(* Logix 5000 project; controller TFF vendor 1 type 14 code 107 rev 34.11; software revision 34.03; part 5 of 36 *)

        [11].DelayTimerSP := 1, [11].ActiveStateCFg := 1, [11].RealInputCfg := 1, [11].InputAddressCfg := 11, [12].Tag := 'XS012', [12].DelayTimer.PRE := 1000, [12].DelayTimerSP := 1, [12].EnableCfg := 1, [12].ActiveStateCFg := 1, [12].RealInputCfg := 1, [12].InputAddressCfg := 12, [13].Tag := 'XC102_3DF', [13].AlarmCurrentValue := 1, [13].Override := 1, [13].DelayTimer.PRE := 1000, [13].DelayTimer.ACC := 1007, [13].DelayTimer.EN := 1, [13].DelayTimer.DN := 1, [13].DelayTimerSP := 1, [13].Priority := 1, [13].EnableCfg := 1, [13].ActiveStateCFg := 1, [13].RealInputCfg := 1, [13].InputAddressCfg := 13, [13].AlarmCfg := 1, [13].OverrideCfg := 1, [13].PriorityCfg := 1, [14].Tag := 'SIC003DF', [14].AlarmCurrentValue := 1, [14].Override := 1, [14].DelayTimer.PRE := 1000, [14].DelayTimer.ACC := 1005, [14].DelayTimer.EN := 1, [14].DelayTimer.DN := 1, [14].DelayTimerSP := 1, [14].Priority := 1, [14].EnableCfg := 1, [14].ActiveStateCFg := 1, [14].RealInputCfg := 1, [14].InputAddressCfg := 14, [14].AlarmCfg := 1, [14].OverrideCfg := 1, [14].PriorityCfg := 1, [15].Tag := 'SRL001', [15].SoftInput := 1, [15].DelayTimer.PRE := 2000, [15].DelayTimerSP := 2, [15].EnableCfg := 1, [15].ActiveStateCFg := 1, [15].RealInputCfg := 1, [15].InputAddressCfg := 15, [16].AlarmCurrentValue := 1, [16].Override := 1, [16].SoftInput := 1, [16].DelayTimer.PRE := 1000, [16].DelayTimer.ACC := 1018, [16].DelayTimer.EN := 1, [16].DelayTimer.DN := 1, [16].DelayTimerSP := 1, [16].Priority := 1,
        [16].ActiveStateCFg := 1, [16].RealInputCfg := 1, [16].InputAddressCfg := 16, [16].OverrideCfg := 1, [16].PriorityCfg := 1, [17].AlarmCurrentValue := 1, [17].Override := 1, [17].SoftInput := 1, [17].DelayTimer.PRE := 1000, [17].DelayTimer.ACC := 1018, [17].DelayTimer.EN := 1, [17].DelayTimer.DN := 1, [17].DelayTimerSP := 1, [17].Priority := 1, [17].ActiveStateCFg := 1, [17].RealInputCfg := 1, [17].InputAddressCfg := 17, [17].OverrideCfg := 1, [17].PriorityCfg := 1, [18].AlarmCurrentValue := 1, [18].Override := 1, [18].DelayTimer.PRE := 1000, [18].DelayTimer.ACC := 1018, [18].DelayTimer.EN := 1, [18].DelayTimer.DN := 1, [18].DelayTimerSP := 1, [18].Priority := 1, [18].ActiveStateCFg := 1, [18].RealInputCfg := 1, [18].InputAddressCfg := 18, [18].OverrideCfg := 1, [18].PriorityCfg := 1, [19].AlarmCurrentValue := 1, [19].Override := 1, [19].DelayTimer.PRE := 1000, [19].DelayTimer.ACC := 1019, [19].DelayTimer.EN := 1, [19].DelayTimer.DN := 1, [19].DelayTimerSP := 1, [19].ActiveStateCFg := 1, [19].RealInputCfg := 1, [19].InputAddressCfg := 19, [19].OverrideCfg := 1, [19].PriorityCfg := 1, [20].AlarmCurrentValue := 1, [20].Override := 1, [20].DelayTimer.PRE := 1000, [20].DelayTimer.ACC := 1019, [20].DelayTimer.EN := 1, [20].DelayTimer.DN := 1, [20].DelayTimerSP := 1, [20].ActiveStateCFg := 1, [20].RealInputCfg := 1, [20].InputAddressCfg := 20, [20].OverrideCfg := 1, [20].PriorityCfg := 1, [21].AlarmCurrentValue := 1, [21].AlarmAck := 1, [21].Alarm := 1, [21].Mimic := 5,
        [21].DelayTimer.PRE := 1000, [21].DelayTimer.ACC := 1003, [21].DelayTimer.EN := 1, [21].DelayTimer.DN := 1, [21].DelayTimerSP := 1, [21].Priority := 1, [21].ActiveStateCFg := 1, [21].RealInputCfg := 1, [21].InputAddressCfg := 21, [21].AlarmONS := 1, [22].AlarmCurrentValue := 1, [22].AlarmAck := 1, [22].Alarm := 1, [22].Mimic := 5, [22].DelayTimer.PRE := 1000, [22].DelayTimer.ACC := 1004, [22].DelayTimer.EN := 1, [22].DelayTimer.DN := 1, [22].DelayTimerSP := 1, [22].Priority := 1, [22].ActiveStateCFg := 1, [22].RealInputCfg := 1, [22].InputAddressCfg := 22, [22].AlarmONS := 1, [23].AlarmCurrentValue := 1, [23].Override := 1, [23].DelayTimer.PRE := 1000, [23].DelayTimer.ACC := 1018, [23].DelayTimer.EN := 1, [23].DelayTimer.DN := 1, [23].DelayTimerSP := 1, [23].Priority := 1, [23].ActiveStateCFg := 1, [23].RealInputCfg := 1, [23].InputAddressCfg := 23, [23].OverrideCfg := 1, [23].PriorityCfg := 1, [24].AlarmCurrentValue := 1, [24].Override := 1, [24].DelayTimer.PRE := 1000, [24].DelayTimer.ACC := 1018, [24].DelayTimer.EN := 1, [24].DelayTimer.DN := 1, [24].DelayTimerSP := 1, [24].Priority := 1, [24].ActiveStateCFg := 1, [24].RealInputCfg := 1, [24].InputAddressCfg := 24, [24].OverrideCfg := 1, [24].PriorityCfg := 1, [25].AlarmCurrentValue := 1, [25].Override := 1, [25].DelayTimer.PRE := 20000, [25].DelayTimerSP := 2, [25].Priority := 1, [25].ActiveStateCFg := 1, [25].RealInputCfg := 1, [25].InputAddressCfg := 25, [25].OverrideCfg := 1, [25].PriorityCfg := 1,
        [25].Cond1Cfg := 1, [27].SoftInput := 1, [28].SoftInput := 1, [29].SoftInput := 1, [30].SoftInput := 1, [34].Tag := 'DI1', [34].Override := 1, [34].SoftInput := 1, [34].ActiveStateCFg := 1, [34].RealInputCfg := 1, [34].InputAddressCfg := 34, [34].OverrideCfg := 1, [34].PriorityCfg := 1, [35].Tag := 'DI2', [35].Override := 1, [35].ActiveStateCFg := 1, [35].RealInputCfg := 1, [35].InputAddressCfg := 35, [35].OverrideCfg := 1, [35].PriorityCfg := 1, [36].Tag := 'DI3', [36].Override := 1, [36].SoftInput := 1, [36].ActiveStateCFg := 1, [36].RealInputCfg := 1, [36].InputAddressCfg := 36, [36].OverrideCfg := 1, [36].PriorityCfg := 1, [37].Tag := 'DI4', [37].Override := 1, [37].ActiveStateCFg := 1, [37].RealInputCfg := 1, [37].InputAddressCfg := 37, [37].OverrideCfg := 1, [37].PriorityCfg := 1, [38].Tag := 'DI5', [38].Override := 1, [38].ActiveStateCFg := 1, [38].RealInputCfg := 1, [38].InputAddressCfg := 38, [38].OverrideCfg := 1, [38].PriorityCfg := 1, [39].Tag := 'DI6', [39].Override := 1, [39].SoftInput := 1, [39].ActiveStateCFg := 1, [39].RealInputCfg := 1, [39].InputAddressCfg := 39, [39].OverrideCfg := 1, [39].PriorityCfg := 1, [40].Tag := 'DI7', [40].Override := 1, [40].ActiveStateCFg := 1, [40].RealInputCfg := 1, [40].InputAddressCfg := 40, [40].OverrideCfg := 1, [40].PriorityCfg := 1, [41].Tag := 'DI8', [41].Override := 1, [41].SoftInput := 1,
        [41].ActiveStateCFg := 1, [41].RealInputCfg := 1, [41].InputAddressCfg := 41, [41].OverrideCfg := 1, [41].PriorityCfg := 1, [50].Tag := 'YA01', [50].AlarmCurrentValue := 1, [50].Alarm := 1, [50].Mimic := 2, [50].SoftInput := 1, [50].Condition1 := 1, [50].DelayTimer.PRE := 60000, [50].DelayTimer.ACC := 60037, [50].DelayTimer.EN := 1, [50].DelayTimer.DN := 1, [50].DelayTimerSP := 60, [50].EnableCfg := 1, [50].InputAddressCfg := 50, [50].AlarmCfg := 1, [50].AlarmStateCfg := 1, [50].OverrideCfg := 1, [50].PriorityCfg := 1, [50].Cond1Cfg := 1, [50].AlarmONS := 1, [51].Tag := 'YA02', [51].AlarmCurrentValue := 1, [51].Alarm := 1, [51].Mimic := 2, [51].SoftInput := 1, [51].Condition1 := 1, [51].DelayTimer.PRE := 60000, [51].DelayTimer.ACC := 60003, [51].DelayTimer.EN := 1, [51].DelayTimer.DN := 1, [51].DelayTimerSP := 60, [51].EnableCfg := 1, [51].InputAddressCfg := 51, [51].AlarmCfg := 1, [51].AlarmStateCfg := 1, [51].OverrideCfg := 1, [51].PriorityCfg := 1, [51].Cond1Cfg := 1, [51].AlarmONS := 1, [52].Tag := 'YA03', [52].AlarmCurrentValue := 1, [52].Alarm := 1, [52].Mimic := 2, [52].SoftInput := 1, [52].Condition1 := 1, [52].DelayTimer.PRE := 60000, [52].DelayTimer.ACC := 60042, [52].DelayTimer.EN := 1, [52].DelayTimer.DN := 1, [52].DelayTimerSP := 60, [52].EnableCfg := 1, [52].InputAddressCfg := 52, [52].AlarmCfg := 1, [52].AlarmStateCfg := 1, [52].OverrideCfg := 1, [52].PriorityCfg := 1,
        [52].Cond1Cfg := 1, [52].AlarmONS := 1, [53].Tag := 'YA04', [53].DelayTimer.PRE := 60000, [53].DelayTimerSP := 60, [53].EnableCfg := 1, [53].ActiveStateCFg := 1, [53].InputAddressCfg := 53, [53].AlarmCfg := 1, [53].AlarmStateCfg := 1, [53].OverrideCfg := 1, [53].PriorityCfg := 1, [54].Tag := 'YA05', [54].DelayTimer.PRE := 60000, [54].DelayTimerSP := 60, [54].EnableCfg := 1, [54].ActiveStateCFg := 1, [54].InputAddressCfg := 54, [54].AlarmCfg := 1, [54].AlarmStateCfg := 1, [54].OverrideCfg := 1, [54].PriorityCfg := 1, [55].Tag := 'YA06', [55].DelayTimer.PRE := 5000, [55].DelayTimerSP := 5, [55].EnableCfg := 1, [55].ActiveStateCFg := 1, [55].InputAddressCfg := 55, [55].AlarmCfg := 1, [55].AlarmStateCfg := 1, [55].OverrideCfg := 1, [55].PriorityCfg := 1, [56].Tag := 'YA07', [56].DelayTimer.PRE := 2000, [56].DelayTimerSP := 2, [56].EnableCfg := 1, [56].ActiveStateCFg := 1, [56].InputAddressCfg := 56, [56].AlarmCfg := 1, [56].AlarmStateCfg := 1, [56].OverrideCfg := 1, [56].PriorityCfg := 1, [57].Tag := 'YA08', [57].DelayTimer.PRE := 5000, [57].DelayTimerSP := 5, [57].Priority := 1, [57].EnableCfg := 1, [57].ActiveStateCFg := 1, [57].InputAddressCfg := 57, [57].AlarmCfg := 1, [57].AlarmStateCfg := 1, [57].OverrideCfg := 1, [57].PriorityCfg := 1, [58].Tag := 'YA09', [58].DelayTimer.PRE := 2000, [58].DelayTimerSP := 2, [58].EnableCfg := 1, [58].ActiveStateCFg := 1, [58].InputAddressCfg := 58, [58].AlarmCfg := 1,
        [58].AlarmStateCfg := 1, [58].OverrideCfg := 1, [58].PriorityCfg := 1, [59].Tag := 'YA10', [59].CurrentValue := 1, [59].Mimic := 1, [59].Priority := 1, [59].EnableCfg := 1, [59].InputAddressCfg := 59, [59].AlarmCfg := 1, [59].AlarmStateCfg := 1, [60].Tag := 'YA11', [60].Override := 1, [60].DelayTimer.PRE := 5000, [60].DelayTimerSP := 5, [60].EnableCfg := 1, [60].ActiveStateCFg := 1, [60].InputAddressCfg := 60, [60].AlarmCfg := 1, [60].AlarmStateCfg := 1, [60].OverrideCfg := 1, [60].PriorityCfg := 1, [61].Tag := 'YA12', [61].Override := 1, [61].EnableCfg := 1, [61].ActiveStateCFg := 1, [61].InputAddressCfg := 61, [61].AlarmCfg := 1, [61].AlarmStateCfg := 1, [61].OverrideCfg := 1, [61].PriorityCfg := 1, [62].Tag := 'YA13', [62].Override := 1, [62].DelayTimer.PRE := 2000, [62].DelayTimerSP := 2, [62].EnableCfg := 1, [62].ActiveStateCFg := 1, [62].InputAddressCfg := 62, [62].AlarmCfg := 1, [62].AlarmStateCfg := 1, [62].OverrideCfg := 1, [62].PriorityCfg := 1, [63].Tag := 'YA14', [63].CurrentValue := 1, [63].Mimic := 1, [63].DelayTimer.PRE := 60000, [63].DelayTimerSP := 60, [63].EnableCfg := 1, [63].InputAddressCfg := 63, [63].AlarmCfg := 1, [63].AlarmStateCfg := 1, [64].Tag := 'UserNCr1', [64].CurrentValue := 1, [64].Mimic := 1, [64].EnableCfg := 1, [64].InputAddressCfg := 64, [65].Tag := 'UserCr1', [65].CurrentValue := 1, [65].Mimic := 1, [65].Priority := 1,
        [65].EnableCfg := 1, [65].InputAddressCfg := 65, [66].Tag := 'UserNCr2', [66].CurrentValue := 1, [66].Mimic := 1, [66].DelayTimer.PRE := 2000, [66].DelayTimerSP := 2, [66].EnableCfg := 1, [66].InputAddressCfg := 66, [67].Tag := 'UserCr2', [67].CurrentValue := 1, [67].Mimic := 1, [67].DelayTimer.PRE := 2000, [67].DelayTimerSP := 2, [67].Priority := 1, [67].EnableCfg := 1, [67].InputAddressCfg := 67, [68].Tag := 'ZSDF', [68].CurrentValue := 1, [68].AlarmCurrentValue := 1, [68].Override := 1, [68].Mimic := 1, [68].SoftInput := 1, [68].DelayTimer.PRE := 1000, [68].DelayTimer.ACC := 1009, [68].DelayTimer.EN := 1, [68].DelayTimer.DN := 1, [68].DelayTimerSP := 1, [68].Priority := 1, [68].EnableCfg := 1, [68].ActiveStateCFg := 1, [68].InputAddressCfg := 68, [68].AlarmCfg := 1, [68].AlarmStateCfg := 1, [68].OverrideCfg := 1, [68].PriorityCfg := 1, [69].Tag := 'YA15', [69].DelayTimer.PRE := 5000, [69].DelayTimerSP := 5, [69].Priority := 1, [69].EnableCfg := 1, [69].ActiveStateCFg := 1, [69].InputAddressCfg := 69, [69].AlarmCfg := 1, [69].AlarmStateCfg := 1, [69].OverrideCfg := 1, [69].PriorityCfg := 1, [70].Tag := 'YA16', [70].DelayTimer.PRE := 2000, [70].DelayTimerSP := 2, [70].EnableCfg := 1, [70].ActiveStateCFg := 1, [70].InputAddressCfg := 70, [70].AlarmCfg := 1, [70].AlarmStateCfg := 1, [70].OverrideCfg := 1, [70].PriorityCfg := 1, [71].Tag := 'YA17', [71].DelayTimer.PRE := 5000, [71].DelayTimerSP := 5,
        [71].Priority := 1, [71].EnableCfg := 1, [71].ActiveStateCFg := 1, [71].InputAddressCfg := 71, [71].AlarmCfg := 1, [71].AlarmStateCfg := 1, [71].OverrideCfg := 1, [71].PriorityCfg := 1, [72].Tag := 'YA18', [72].DelayTimer.PRE := 2000, [72].DelayTimerSP := 2, [72].EnableCfg := 1, [72].ActiveStateCFg := 1, [72].InputAddressCfg := 72, [72].AlarmCfg := 1, [72].AlarmStateCfg := 1, [72].OverrideCfg := 1, [72].PriorityCfg := 1, [73].Tag := 'YA19', [73].DelayTimer.PRE := 5000, [73].DelayTimerSP := 5, [73].Priority := 1, [73].EnableCfg := 1, [73].ActiveStateCFg := 1, [73].InputAddressCfg := 73, [73].AlarmCfg := 1, [73].AlarmStateCfg := 1, [73].OverrideCfg := 1, [73].PriorityCfg := 1, [74].Tag := 'YA20', [74].DelayTimer.PRE := 2000, [74].DelayTimerSP := 2, [74].EnableCfg := 1, [74].ActiveStateCFg := 1, [74].InputAddressCfg := 74, [74].AlarmCfg := 1, [74].AlarmStateCfg := 1, [74].OverrideCfg := 1, [74].PriorityCfg := 1, [75].Tag := 'YA21', [75].DelayTimer.PRE := 5000, [75].DelayTimerSP := 5, [75].Priority := 1, [75].EnableCfg := 1, [75].ActiveStateCFg := 1, [75].InputAddressCfg := 75, [75].AlarmCfg := 1, [75].AlarmStateCfg := 1, [75].OverrideCfg := 1, [75].PriorityCfg := 1, [76].Tag := 'YA22', [76].DelayTimer.PRE := 5000, [76].DelayTimerSP := 5, [76].Priority := 1, [76].ActiveStateCFg := 1, [76].InputAddressCfg := 76, [76].AlarmStateCfg := 1, [76].OverrideCfg := 1, [76].PriorityCfg := 1, [77].Override := 1,
        [77].DelayTimer.PRE := 2000, [77].DelayTimerSP := 2, [77].EnableCfg := 1, [77].ActiveStateCFg := 1, [77].InputAddressCfg := 77, [77].AlarmCfg := 1, [77].AlarmStateCfg := 1, [77].OverrideCfg := 1, [78].CurrentValue := 1, [78].AlarmCurrentValue := 1, [78].AlarmAck := 1, [78].Alarm := 1, [78].Mimic := 5, [78].SoftInput := 1, [78].DelayTimer.ACC := 45, [78].DelayTimer.EN := 1, [78].DelayTimer.DN := 1, [78].DelayTimerSP := 2, [78].AlarmONS := 1, [79].CurrentValue := 1, [79].AlarmCurrentValue := 1, [79].Mimic := 1, [79].DelayTimer.ACC := 44, [79].DelayTimer.EN := 1, [79].DelayTimer.DN := 1, [79].DelayTimerSP := 2, [80].CurrentValue := 1, [80].AlarmCurrentValue := 1, [80].Mimic := 1, [80].DelayTimer.ACC := 44, [80].DelayTimer.EN := 1, [80].DelayTimer.DN := 1, [80].DelayTimerSP := 2, [81].CurrentValue := 1, [81].AlarmCurrentValue := 1, [81].Mimic := 1, [81].DelayTimer.ACC := 44, [81].DelayTimer.EN := 1, [81].DelayTimer.DN := 1, [81].DelayTimerSP := 2, [82].CurrentValue := 1, [82].AlarmCurrentValue := 1, [82].Mimic := 1, [82].DelayTimer.ACC := 44, [82].DelayTimer.EN := 1, [82].DelayTimer.DN := 1, [82].DelayTimerSP := 2, [83].CurrentValue := 1, [83].AlarmCurrentValue := 1, [83].AlarmAck := 1, [83].Alarm := 1, [83].Mimic := 5, [83].SoftInput := 1, [83].DelayTimer.ACC := 44, [83].DelayTimer.EN := 1, [83].DelayTimer.DN := 1, [83].DelayTimerSP := 2, [83].AlarmONS := 1, [84].CurrentValue := 1, [84].Mimic := 1,
        [84].DelayTimerSP := 2, [85].CurrentValue := 1, [85].AlarmCurrentValue := 1, [85].AlarmAck := 1, [85].Alarm := 1, [85].Mimic := 3, [85].SoftInput := 1, [85].DelayTimer.ACC := 2021, [85].DelayTimer.EN := 1, [85].DelayTimer.DN := 1, [85].DelayTimerSP := 2, [85].AlarmONS := 1, [86].CurrentValue := 1, [86].Mimic := 1, [86].DelayTimerSP := 2, [87].CurrentValue := 1, [87].Mimic := 1, [87].DelayTimerSP := 2, [88].CurrentValue := 1, [88].Mimic := 1, [88].DelayTimerSP := 2, [89].CurrentValue := 1, [89].Mimic := 1, [89].DelayTimerSP := 2, [90].Tag := 'AI101_SIG', [90].Override := 1, [90].DelayTimer.PRE := 2000, [90].DelayTimerSP := 2, [90].Priority := 1, [90].EnableCfg := 1, [90].ActiveStateCFg := 1, [90].InputAddressCfg := 90, [90].AlarmCfg := 1, [90].AlarmStateCfg := 1, [90].OverrideCfg := 1, [90].PriorityCfg := 1, [91].Tag := 'AI102_SIG', [91].Override := 1, [91].DelayTimer.PRE := 2000, [91].DelayTimerSP := 2, [91].Priority := 1, [91].EnableCfg := 1, [91].ActiveStateCFg := 1, [91].InputAddressCfg := 91, [91].AlarmCfg := 1, [91].AlarmStateCfg := 1, [91].OverrideCfg := 1, [91].PriorityCfg := 1, [92].Tag := 'AI103_SIG', [92].Override := 1, [92].DelayTimer.PRE := 2000, [92].DelayTimerSP := 2, [92].Priority := 1, [92].EnableCfg := 1, [92].ActiveStateCFg := 1, [92].InputAddressCfg := 92, [92].AlarmCfg := 1, [92].AlarmStateCfg := 1, [92].OverrideCfg := 1, [92].PriorityCfg := 1,
        [93].Tag := 'FI101_SIG', [93].CurrentValue := 1, [93].AlarmCurrentValue := 1, [93].Override := 1, [93].Mimic := 1, [93].DelayTimer.PRE := 5000, [93].DelayTimer.ACC := 5039, [93].DelayTimer.EN := 1, [93].DelayTimer.DN := 1, [93].DelayTimerSP := 5, [93].ActiveStateCFg := 1, [93].InputAddressCfg := 93, [93].AlarmStateCfg := 1, [93].OverrideCfg := 1, [93].PriorityCfg := 1, [94].Tag := 'WI001_SIG', [94].Override := 1, [94].DelayTimer.PRE := 2000, [94].DelayTimerSP := 2, [94].Priority := 1, [94].EnableCfg := 1, [94].ActiveStateCFg := 1, [94].InputAddressCfg := 94, [94].AlarmCfg := 1, [94].AlarmStateCfg := 1, [94].OverrideCfg := 1, [94].PriorityCfg := 1, [95].Tag := 'WI101_SIG', [95].DelayTimer.PRE := 2000, [95].DelayTimerSP := 2, [95].Priority := 1, [95].ActiveStateCFg := 1, [95].InputAddressCfg := 95, [95].AlarmStateCfg := 1, [95].OverrideCfg := 1, [95].PriorityCfg := 1, [96].Tag := 'WI102_SIG', [96].CurrentValue := 1, [96].AlarmCurrentValue := 1, [96].Override := 1, [96].Mimic := 1, [96].SoftInput := 1, [96].DelayTimer.PRE := 2000, [96].DelayTimer.ACC := 4082459, [96].DelayTimer.EN := 1, [96].DelayTimer.DN := 1, [96].DelayTimerSP := 2, [96].EnableCfg := 1, [96].ActiveStateCFg := 1, [96].InputAddressCfg := 96, [96].AlarmCfg := 1, [96].AlarmStateCfg := 1, [96].OverrideCfg := 1, [96].PriorityCfg := 1, [97].Tag := 'PI001_SIG', [97].Override := 1, [97].DelayTimer.PRE := 2000, [97].DelayTimerSP := 2, [97].Priority := 1, [97].EnableCfg := 1,
        [97].ActiveStateCFg := 1, [97].InputAddressCfg := 97, [97].AlarmCfg := 1, [97].AlarmStateCfg := 1, [97].OverrideCfg := 1, [97].PriorityCfg := 1, [98].Tag := 'PI002_SIG', [98].Override := 1, [98].DelayTimer.PRE := 2000, [98].DelayTimerSP := 2, [98].Priority := 1, [98].EnableCfg := 1, [98].ActiveStateCFg := 1, [98].InputAddressCfg := 98, [98].AlarmCfg := 1, [98].AlarmStateCfg := 1, [98].OverrideCfg := 1, [98].PriorityCfg := 1, [99].Tag := 'PI101_SIG', [99].Override := 1, [99].DelayTimer.PRE := 2000, [99].DelayTimerSP := 2, [99].Priority := 1, [99].EnableCfg := 1, [99].ActiveStateCFg := 1, [99].InputAddressCfg := 99, [99].AlarmCfg := 1, [99].AlarmStateCfg := 1, [99].OverrideCfg := 1, [99].PriorityCfg := 1, [100].Tag := 'PI401_SIG', [100].Override := 1, [100].DelayTimer.PRE := 2000, [100].DelayTimerSP := 2, [100].Priority := 1, [100].EnableCfg := 1, [100].ActiveStateCFg := 1, [100].InputAddressCfg := 100, [100].AlarmCfg := 1, [100].AlarmStateCfg := 1, [100].OverrideCfg := 1, [100].PriorityCfg := 1, [101].Tag := 'TI001_SIG', [101].Override := 1, [101].DelayTimer.PRE := 2000, [101].DelayTimerSP := 2, [101].Priority := 1, [101].EnableCfg := 1, [101].ActiveStateCFg := 1, [101].InputAddressCfg := 101, [101].AlarmCfg := 1, [101].AlarmStateCfg := 1, [101].OverrideCfg := 1, [101].PriorityCfg := 1, [102].Tag := 'PCV001_SIG', [102].Override := 1, [102].DelayTimer.PRE := 2000, [102].DelayTimerSP := 2, [102].Priority := 1, [102].EnableCfg := 1,
        [102].ActiveStateCFg := 1, [102].InputAddressCfg := 102, [102].AlarmCfg := 1, [102].AlarmStateCfg := 1, [102].OverrideCfg := 1, [102].PriorityCfg := 1, [103].Tag := 'PCV101_SIG', [103].Override := 1, [103].DelayTimer.PRE := 2000, [103].DelayTimerSP := 2, [103].Priority := 1, [103].EnableCfg := 1, [103].ActiveStateCFg := 1, [103].InputAddressCfg := 103, [103].AlarmCfg := 1, [103].AlarmStateCfg := 1, [103].OverrideCfg := 1, [103].PriorityCfg := 1, [104].Tag := 'MIX001_SIG', [104].Override := 1, [104].DelayTimer.PRE := 2000, [104].DelayTimerSP := 2, [104].Priority := 1, [104].EnableCfg := 1, [104].ActiveStateCFg := 1, [104].InputAddressCfg := 104, [104].AlarmCfg := 1, [104].AlarmStateCfg := 1, [104].OverrideCfg := 1, [104].PriorityCfg := 1, [105].Tag := 'AI104_SIG', [105].CurrentValue := 1, [105].AlarmCurrentValue := 1, [105].Mimic := 1, [105].SoftInput := 1, [105].DelayTimer.PRE := 2000, [105].DelayTimer.ACC := 47, [105].DelayTimer.EN := 1, [105].DelayTimer.DN := 1, [105].DelayTimerSP := 2, [105].Priority := 1, [105].ActiveStateCFg := 1, [105].InputAddressCfg := 105, [105].AlarmStateCfg := 1, [105].OverrideCfg := 1, [105].PriorityCfg := 1, [106].ActiveStateCFg := 1, [106].InputAddressCfg := 106, [106].AlarmStateCfg := 1, [106].OverrideCfg := 1, [106].PriorityCfg := 1);   // Digital Point Array
        [94]   // Feed Bag Weight Signal Default
        [95]   // Filtrate Weight Signal Default
        [100]   // Transfer Pump Pressure Signal Default
        [52]   // Historical Data collection failure
        [96]   // Customer Filtrate Weight Signal Default
        [102]   // PCV001 Position Signal Default
        [101]   // Feed Bag Temperature Signal Default
        [103]   // PCV101 Position Signal Default
        [99]   // Filtrate Pressure Signal Default
        [51]   // CCP Runtime communication failure
        [69]   // YA15 Node 3 Communication Failure
        [90]   // Filtrate Conductivity Signal Default
        [71]   // YA17 Node 4 Communication Failure
        [73]   // YA19 Node 5 Communication Failure
        [75]   // YA21 IND331 Communication Failure
        [76]   // YA22 IND131 Communication Failure
        [106]   // Retentate Flow Signal Default
        [15]   // Tank Skid Remote / Standalone
        [68]   // ZSDF Clamshell Locking Defect
        [11]   // Pump P001 Type
        [12]   // Pump P002 Type
        [53]   // Hard Drive Overload
        [54]   // Database Overload
        [8]   // Feed Pump Defect
        [50]   // PC to PLC communication failure
        [98]   // Rentate Pressure Signal Default
        [59]   // PLC Program Major Fault
        [104]   // Mixer Speed Signal Default
        [105]   // Filtrate pH Signal Default
        [60]   // Database Corrupted
        [55]   // Node 0 communication failure
        [57]   // Node 1 communication failure
        [1]   // Door Closed
        [62]   // Tank Size Mismatch
        [9]   // Transfer Pump Defect
        [63]   // SQL Server Write Failure
        [5]   // Transfer Pump High Pressure
        [64]   // User Non Critical Alarm 1
        [77]   // YA41 Operating Time Exceeded
        [6]   // Clamshell Locking 1 Closed
        [7]   // Clamshell Locking 2 Closed
        [93]   // Filtrate Flow Signal Default
        [97]   // Feed Pressure Signal Default
        [66]   // User Non Critical Alarm 2
        [13]   // C8000 Defect
        [14]   // Mixer Defect
        [3]   // Emergency Stop
        [10]   // Manifold Valves Air Defect
        [2]   // Door to Frame Locking Defect
        [91]   // Filtrate UV Signal Default
        [56]   // Node 0 internal defect
        [58]   // Node 1 internal defect
        [4]   // Feed Pump High Pressure
        [61]   // Unauthorized Accesses
        [65]   // User Critical Alarm 1
        [67]   // User Critical Alarm 2
        [70]   // YA16 Node 3 Internal Defect
        [72]   // YA18 Node 4 Internal Defect
        [74]   // YA20 Node 5 Internal Defect
        [92]   // Filtrate UV Signal Default
        [0]   // Valves Air Defect
   DigitalPoint_Storage : DigitalPoint[6,150] := ([0,0].Tag := 'PISL601', [0,0].AlarmCurrentValue := 1, [0,0].AlarmAck := 1, [0,0].Alarm := 1, [0,0].Mimic := 5, [0,0].DelayTimer.PRE := 2000, [0,0].DelayTimer.ACC := 2025, [0,0].DelayTimer.EN := 1, [0,0].DelayTimer.DN := 1, [0,0].DelayTimerSP := 2, [0,0].Priority := 1, [0,0].EnableCfg := 1, [0,0].ActiveStateCFg := 1, [0,0].RealInputCfg := 1, [0,0].AlarmCfg := 1, [0,0].OverrideCfg := 1, [0,0].PriorityCfg := 1, [0,0].AlarmONS := 1, [0,1].Tag := 'PISL602', [0,1].AlarmCurrentValue := 1, [0,1].AlarmAck := 1, [0,1].Alarm := 1, [0,1].Mimic := 5, [0,1].Condition2 := 1, [0,1].DelayTimer.PRE := 2000, [0,1].DelayTimer.ACC := 2053, [0,1].DelayTimer.EN := 1, [0,1].DelayTimer.DN := 1, [0,1].DelayTimerSP := 2, [0,1].Priority := 1, [0,1].EnableCfg := 1, [0,1].ActiveStateCFg := 1, [0,1].RealInputCfg := 1, [0,1].InputAddressCfg := 1, [0,1].AlarmCfg := 1, [0,1].OverrideCfg := 1, [0,1].PriorityCfg := 1, [0,1].AlarmONS := 1, [0,2].Tag := 'ES001', [0,2].AlarmCurrentValue := 1, [0,2].AlarmAck := 1, [0,2].Alarm := 1, [0,2].Mimic := 5, [0,2].DelayTimer.PRE := 1000, [0,2].DelayTimer.ACC := 1047, [0,2].DelayTimer.EN := 1, [0,2].DelayTimer.DN := 1, [0,2].DelayTimerSP := 1, [0,2].Priority := 1, [0,2].EnableCfg := 1, [0,2].ActiveStateCFg := 1, [0,2].RealInputCfg := 1, [0,2].InputAddressCfg := 2, [0,2].AlarmCfg := 1, [0,2].AlarmONS := 1, [0,3].Tag := 'RSBUZZ', [0,3].DelayTimer.PRE := 2000, [0,3].DelayTimerSP := 2, [0,3].EnableCfg := 1, [0,3].ActiveStateCFg := 1,
        [0,3].RealInputCfg := 1, [0,3].InputAddressCfg := 3, [0,4].Tag := 'DF24VDC', [0,4].AlarmCurrentValue := 1, [0,4].AlarmAck := 1, [0,4].Alarm := 1, [0,4].Mimic := 5, [0,4].DelayTimer.PRE := 1000, [0,4].DelayTimer.ACC := 1048, [0,4].DelayTimer.EN := 1, [0,4].DelayTimer.DN := 1, [0,4].DelayTimerSP := 1, [0,4].Priority := 1, [0,4].EnableCfg := 1, [0,4].ActiveStateCFg := 1, [0,4].RealInputCfg := 1, [0,4].InputAddressCfg := 4, [0,4].AlarmCfg := 1, [0,4].OverrideCfg := 1, [0,4].PriorityCfg := 1, [0,4].AlarmONS := 1, [0,5].Tag := 'ZS008', [0,5].AlarmCurrentValue := 1, [0,5].AlarmAck := 1, [0,5].Alarm := 1, [0,5].Mimic := 5, [0,5].DelayTimer.PRE := 1000, [0,5].DelayTimer.ACC := 1048, [0,5].DelayTimer.EN := 1, [0,5].DelayTimer.DN := 1, [0,5].DelayTimerSP := 1, [0,5].Priority := 1, [0,5].EnableCfg := 1, [0,5].ActiveStateCFg := 1, [0,5].RealInputCfg := 1, [0,5].InputAddressCfg := 5, [0,5].AlarmCfg := 1, [0,5].OverrideCfg := 1, [0,5].AlarmONS := 1, [0,6].Tag := 'ZS001', [0,6].DelayTimer.PRE := 2000, [0,6].DelayTimerSP := 2, [0,6].EnableCfg := 1, [0,6].ActiveStateCFg := 1, [0,6].RealInputCfg := 1, [0,6].InputAddressCfg := 6, [0,7].Tag := 'ZS002', [0,7].DelayTimer.PRE := 2000, [0,7].DelayTimerSP := 2, [0,7].EnableCfg := 1, [0,7].ActiveStateCFg := 1, [0,7].RealInputCfg := 1, [0,7].InputAddressCfg := 7, [0,8].Tag := 'ZS003', [0,8].DelayTimer.PRE := 2000, [0,8].DelayTimerSP := 2, [0,8].EnableCfg := 1, [0,8].ActiveStateCFg := 1, [0,8].RealInputCfg := 1, [0,8].InputAddressCfg := 8,
        [0,9].Tag := 'ZS004', [0,9].DelayTimer.PRE := 2000, [0,9].DelayTimerSP := 2, [0,9].EnableCfg := 1, [0,9].ActiveStateCFg := 1, [0,9].RealInputCfg := 1, [0,9].InputAddressCfg := 9, [0,10].Tag := 'ZS005', [0,10].DelayTimer.PRE := 2000, [0,10].DelayTimerSP := 2, [0,10].EnableCfg := 1, [0,10].ActiveStateCFg := 1, [0,10].RealInputCfg := 1, [0,10].InputAddressCfg := 10, [0,11].Tag := 'ZS006', [0,11].DelayTimer.PRE := 2000, [0,11].DelayTimerSP := 2, [0,11].EnableCfg := 1, [0,11].ActiveStateCFg := 1, [0,11].RealInputCfg := 1, [0,11].InputAddressCfg := 11, [0,12].Tag := 'ZS007', [0,12].DelayTimer.PRE := 2000, [0,12].DelayTimerSP := 2, [0,12].EnableCfg := 1, [0,12].ActiveStateCFg := 1, [0,12].RealInputCfg := 1, [0,12].InputAddressCfg := 12, [0,13].Tag := 'ZS008', [0,13].AlarmCurrentValue := 1, [0,13].DelayTimer.PRE := 20000, [0,13].DelayTimerSP := 2, [0,13].Priority := 1, [0,13].EnableCfg := 1, [0,13].ActiveStateCFg := 1, [0,13].RealInputCfg := 1, [0,13].InputAddressCfg := 13, [0,13].AlarmCfg := 1, [0,13].OverrideCfg := 1, [0,13].PriorityCfg := 1, [0,13].Cond1Cfg := 1, [0,14].Tag := 'XS011', [0,14].DelayTimer.PRE := 2000, [0,14].DelayTimerSP := 2, [0,14].EnableCfg := 1, [0,14].ActiveStateCFg := 1, [0,14].RealInputCfg := 1, [0,14].InputAddressCfg := 14, [0,15].Tag := 'XS012', [0,15].SoftInput := 1, [0,15].DelayTimer.PRE := 2000, [0,15].DelayTimerSP := 2, [0,15].EnableCfg := 1, [0,15].ActiveStateCFg := 1, [0,15].RealInputCfg := 1, [0,15].InputAddressCfg := 15, [0,16].Tag := 'SIC001DF', [0,16].AlarmCurrentValue := 1, [0,16].AlarmAck := 1, [0,16].Alarm := 1,
        [0,16].Mimic := 5, [0,16].SoftInput := 1, [0,16].DelayTimer.PRE := 1000, [0,16].DelayTimer.ACC := 1046, [0,16].DelayTimer.EN := 1, [0,16].DelayTimer.DN := 1, [0,16].DelayTimerSP := 1, [0,16].Priority := 1, [0,16].EnableCfg := 1, [0,16].ActiveStateCFg := 1, [0,16].RealInputCfg := 1, [0,16].InputAddressCfg := 16, [0,16].AlarmCfg := 1, [0,16].OverrideCfg := 1, [0,16].PriorityCfg := 1, [0,16].AlarmONS := 1, [0,17].Tag := 'SIC002DF', [0,17].AlarmCurrentValue := 1, [0,17].AlarmAck := 1, [0,17].Alarm := 1, [0,17].Mimic := 5, [0,17].SoftInput := 1, [0,17].DelayTimer.PRE := 1000, [0,17].DelayTimer.ACC := 1046, [0,17].DelayTimer.EN := 1, [0,17].DelayTimer.DN := 1, [0,17].DelayTimerSP := 1, [0,17].Priority := 1, [0,17].EnableCfg := 1, [0,17].ActiveStateCFg := 1, [0,17].RealInputCfg := 1, [0,17].InputAddressCfg := 17, [0,17].AlarmCfg := 1, [0,17].OverrideCfg := 1, [0,17].PriorityCfg := 1, [0,17].AlarmONS := 1, [0,18].Tag := 'AA008', [0,18].AlarmCurrentValue := 1, [0,18].AlarmAck := 1, [0,18].Alarm := 1, [0,18].Mimic := 5, [0,18].DelayTimer.PRE := 1000, [0,18].DelayTimer.ACC := 1046, [0,18].DelayTimer.EN := 1, [0,18].DelayTimer.DN := 1, [0,18].DelayTimerSP := 1, [0,18].Priority := 1, [0,18].EnableCfg := 1, [0,18].ActiveStateCFg := 1, [0,18].RealInputCfg := 1, [0,18].InputAddressCfg := 18, [0,18].AlarmCfg := 1, [0,18].OverrideCfg := 1, [0,18].PriorityCfg := 1, [0,18].AlarmONS := 1, [0,19].Tag := 'LSH001', [0,19].AlarmCurrentValue := 1, [0,19].Override := 1, [0,19].DelayTimer.PRE := 1000, [0,19].DelayTimer.ACC := 1058,
        [0,19].DelayTimer.EN := 1, [0,19].DelayTimer.DN := 1, [0,19].DelayTimerSP := 1, [0,19].EnableCfg := 1, [0,19].ActiveStateCFg := 1, [0,19].RealInputCfg := 1, [0,19].InputAddressCfg := 19, [0,19].AlarmCfg := 1, [0,19].OverrideCfg := 1, [0,19].PriorityCfg := 1, [0,20].Tag := 'LSL002', [0,20].AlarmCurrentValue := 1, [0,20].Override := 1, [0,20].DelayTimer.PRE := 1000, [0,20].DelayTimer.ACC := 1059, [0,20].DelayTimer.EN := 1, [0,20].DelayTimer.DN := 1, [0,20].DelayTimerSP := 1, [0,20].EnableCfg := 1, [0,20].ActiveStateCFg := 1, [0,20].RealInputCfg := 1, [0,20].InputAddressCfg := 20, [0,20].AlarmCfg := 1, [0,20].OverrideCfg := 1, [0,20].PriorityCfg := 1, [0,21].Tag := 'PSH001', [0,21].AlarmCurrentValue := 1, [0,21].AlarmAck := 1, [0,21].Alarm := 1, [0,21].Mimic := 5, [0,21].DelayTimer.PRE := 1000, [0,21].DelayTimer.ACC := 1045, [0,21].DelayTimer.EN := 1, [0,21].DelayTimer.DN := 1, [0,21].DelayTimerSP := 1, [0,21].Priority := 1, [0,21].EnableCfg := 1, [0,21].ActiveStateCFg := 1, [0,21].RealInputCfg := 1, [0,21].InputAddressCfg := 21, [0,21].AlarmCfg := 1, [0,21].AlarmONS := 1, [0,22].Tag := 'PSH002', [0,22].AlarmCurrentValue := 1, [0,22].AlarmAck := 1, [0,22].Alarm := 1, [0,22].Mimic := 5, [0,22].DelayTimer.PRE := 1000, [0,22].DelayTimer.ACC := 1045, [0,22].DelayTimer.EN := 1, [0,22].DelayTimer.DN := 1, [0,22].DelayTimerSP := 1, [0,22].Priority := 1, [0,22].EnableCfg := 1, [0,22].ActiveStateCFg := 1, [0,22].RealInputCfg := 1, [0,22].InputAddressCfg := 22, [0,22].AlarmCfg := 1, [0,22].AlarmONS := 1, [0,23].Tag := 'DF48VP001',
        [0,23].AlarmCurrentValue := 1, [0,23].AlarmAck := 1, [0,23].Alarm := 1, [0,23].Mimic := 5, [0,23].DelayTimer.PRE := 1000, [0,23].DelayTimer.ACC := 1045, [0,23].DelayTimer.EN := 1, [0,23].DelayTimer.DN := 1, [0,23].DelayTimerSP := 1, [0,23].Priority := 1, [0,23].EnableCfg := 1, [0,23].ActiveStateCFg := 1, [0,23].RealInputCfg := 1, [0,23].InputAddressCfg := 23, [0,23].AlarmCfg := 1, [0,23].OverrideCfg := 1, [0,23].PriorityCfg := 1, [0,23].AlarmONS := 1, [0,24].Tag := 'DF48VP002', [0,24].AlarmCurrentValue := 1, [0,24].AlarmAck := 1, [0,24].Alarm := 1, [0,24].Mimic := 5, [0,24].DelayTimer.PRE := 1000, [0,24].DelayTimer.ACC := 1046, [0,24].DelayTimer.EN := 1, [0,24].DelayTimer.DN := 1, [0,24].DelayTimerSP := 1, [0,24].Priority := 1, [0,24].EnableCfg := 1, [0,24].ActiveStateCFg := 1, [0,24].RealInputCfg := 1, [0,24].InputAddressCfg := 24, [0,24].AlarmCfg := 1, [0,24].OverrideCfg := 1, [0,24].PriorityCfg := 1, [0,24].AlarmONS := 1, [0,25].Tag := 'XS002', [0,25].AlarmCurrentValue := 1, [0,25].DelayTimer.PRE := 20000, [0,25].DelayTimerSP := 2, [0,25].Priority := 1, [0,25].EnableCfg := 1, [0,25].ActiveStateCFg := 1, [0,25].RealInputCfg := 1, [0,25].InputAddressCfg := 25, [0,25].AlarmCfg := 1, [0,25].OverrideCfg := 1, [0,25].PriorityCfg := 1, [0,25].Cond1Cfg := 1, [0,26].Override := 1, [0,26].ActiveStateCFg := 1, [0,26].RealInputCfg := 1, [0,26].InputAddressCfg := 26, [0,26].OverrideCfg := 1, [0,26].PriorityCfg := 1, [0,27].Override := 1, [0,27].SoftInput := 1, [0,27].ActiveStateCFg := 1, [0,27].RealInputCfg := 1,
        [0,27].InputAddressCfg := 27, [0,27].OverrideCfg := 1, [0,27].PriorityCfg := 1, [0,28].Override := 1, [0,28].SoftInput := 1, [0,28].ActiveStateCFg := 1, [0,28].RealInputCfg := 1, [0,28].InputAddressCfg := 28, [0,28].OverrideCfg := 1, [0,28].PriorityCfg := 1, [0,29].Override := 1, [0,29].SoftInput := 1, [0,29].ActiveStateCFg := 1, [0,29].RealInputCfg := 1, [0,29].InputAddressCfg := 29, [0,29].OverrideCfg := 1, [0,29].PriorityCfg := 1, [0,30].Override := 1, [0,30].SoftInput := 1, [0,30].ActiveStateCFg := 1, [0,30].RealInputCfg := 1, [0,30].InputAddressCfg := 30, [0,30].OverrideCfg := 1, [0,30].PriorityCfg := 1, [0,31].Override := 1, [0,31].ActiveStateCFg := 1, [0,31].RealInputCfg := 1, [0,31].InputAddressCfg := 31, [0,31].OverrideCfg := 1, [0,31].PriorityCfg := 1, [0,34].Tag := 'DI1', [0,34].Override := 1, [0,34].SoftInput := 1, [0,34].EnableCfg := 1, [0,34].ActiveStateCFg := 1, [0,34].RealInputCfg := 1, [0,34].InputAddressCfg := 34, [0,34].OverrideCfg := 1, [0,34].PriorityCfg := 1, [0,35].Tag := 'DI2', [0,35].Override := 1, [0,35].EnableCfg := 1, [0,35].ActiveStateCFg := 1, [0,35].RealInputCfg := 1, [0,35].InputAddressCfg := 35, [0,35].OverrideCfg := 1, [0,35].PriorityCfg := 1, [0,36].Tag := 'DI3', [0,36].Override := 1, [0,36].SoftInput := 1, [0,36].EnableCfg := 1, [0,36].ActiveStateCFg := 1, [0,36].RealInputCfg := 1, [0,36].InputAddressCfg := 36, [0,36].OverrideCfg := 1, [0,36].PriorityCfg := 1, [0,37].Tag := 'DI4', [0,37].Override := 1, [0,37].EnableCfg := 1, [0,37].ActiveStateCFg := 1,
        [0,37].RealInputCfg := 1, [0,37].InputAddressCfg := 37, [0,37].OverrideCfg := 1, [0,37].PriorityCfg := 1, [0,38].Tag := 'DI5', [0,38].Override := 1, [0,38].EnableCfg := 1, [0,38].ActiveStateCFg := 1, [0,38].RealInputCfg := 1, [0,38].InputAddressCfg := 38, [0,38].OverrideCfg := 1, [0,38].PriorityCfg := 1, [0,39].Tag := 'DI6', [0,39].Override := 1, [0,39].SoftInput := 1, [0,39].EnableCfg := 1, [0,39].ActiveStateCFg := 1, [0,39].RealInputCfg := 1, [0,39].InputAddressCfg := 39, [0,39].OverrideCfg := 1, [0,39].PriorityCfg := 1, [0,40].Tag := 'DI7', [0,40].Override := 1, [0,40].EnableCfg := 1, [0,40].ActiveStateCFg := 1, [0,40].RealInputCfg := 1, [0,40].InputAddressCfg := 40, [0,40].OverrideCfg := 1, [0,40].PriorityCfg := 1, [0,41].Tag := 'DI8', [0,41].Override := 1, [0,41].EnableCfg := 1, [0,41].ActiveStateCFg := 1, [0,41].RealInputCfg := 1, [0,41].InputAddressCfg := 41, [0,41].OverrideCfg := 1, [0,41].PriorityCfg := 1, [0,50].Tag := 'YA01', [0,50].Desc := 'PC to PLC Com. Failure', [0,50].AlarmCurrentValue := 1, [0,50].SoftInput := 1, [0,50].Condition1 := 1, [0,50].Cond1Text := 'HMI HeartBeat received', [0,50].DelayTimer.PRE := 60000, [0,50].DelayTimer.ACC := 442, [0,50].DelayTimer.EN := 1, [0,50].DelayTimer.TT := 1, [0,50].DelayTimerSP := 60, [0,50].EnableCfg := 1, [0,50].InputAddressCfg := 50, [0,50].AlarmCfg := 1, [0,50].AlarmStateCfg := 1, [0,50].OverrideCfg := 1, [0,50].PriorityCfg := 1, [0,50].Cond1Cfg := 1, [0,51].Tag := 'YA02', [0,51].Desc := 'CCP Runtime Com. Failure', [0,51].AlarmCurrentValue := 1, [0,51].Alarm := 1, [0,51].Mimic := 2,
        [0,51].SoftInput := 1, [0,51].Condition1 := 1, [0,51].Cond1Text := 'HMI HeartBeat received', [0,51].DelayTimer.PRE := 60000, [0,51].DelayTimer.ACC := 60061, [0,51].DelayTimer.EN := 1, [0,51].DelayTimer.DN := 1, [0,51].DelayTimerSP := 60, [0,51].EnableCfg := 1, [0,51].InputAddressCfg := 51, [0,51].AlarmCfg := 1, [0,51].AlarmStateCfg := 1, [0,51].OverrideCfg := 1, [0,51].PriorityCfg := 1, [0,51].Cond1Cfg := 1, [0,51].AlarmONS := 1, [0,52].Tag := 'YA03', [0,52].Desc := 'Hist. Data Collect. Fail', [0,52].AlarmCurrentValue := 1, [0,52].Alarm := 1, [0,52].Mimic := 2, [0,52].SoftInput := 1, [0,52].Condition1 := 1, [0,52].Cond1Text := 'HMI HeartBeat received', [0,52].DelayTimer.PRE := 60000, [0,52].DelayTimer.ACC := 1286, [0,52].DelayTimer.EN := 1, [0,52].DelayTimer.TT := 1, [0,52].DelayTimerSP := 60, [0,52].EnableCfg := 1, [0,52].InputAddressCfg := 52, [0,52].AlarmCfg := 1, [0,52].AlarmStateCfg := 1, [0,52].OverrideCfg := 1, [0,52].PriorityCfg := 1, [0,52].Cond1Cfg := 1, [0,52].AlarmONS := 1, [0,53].Tag := 'YA04', [0,53].Desc := 'HDD OverLoad', [0,53].DelayTimer.PRE := 60000, [0,53].DelayTimerSP := 60, [0,53].EnableCfg := 1, [0,53].ActiveStateCFg := 1, [0,53].InputAddressCfg := 53, [0,53].AlarmCfg := 1, [0,53].AlarmStateCfg := 1, [0,53].OverrideCfg := 1, [0,53].PriorityCfg := 1, [0,54].Tag := 'YA05', [0,54].DelayTimer.PRE := 60000, [0,54].DelayTimerSP := 60, [0,54].EnableCfg := 1, [0,54].ActiveStateCFg := 1, [0,54].InputAddressCfg := 54, [0,54].AlarmCfg := 1, [0,54].AlarmStateCfg := 1, [0,54].OverrideCfg := 1, [0,54].PriorityCfg := 1, [0,55].Tag := 'YA06', [0,55].CurrentValue := 1,
        [0,55].AlarmCurrentValue := 1, [0,55].AlarmAck := 1, [0,55].Alarm := 1, [0,55].Mimic := 5, [0,55].SoftInput := 1, [0,55].DelayTimer.PRE := 5000, [0,55].DelayTimer.ACC := 5038, [0,55].DelayTimer.EN := 1, [0,55].DelayTimer.DN := 1, [0,55].DelayTimerSP := 5, [0,55].Priority := 1, [0,55].EnableCfg := 1, [0,55].ActiveStateCFg := 1, [0,55].InputAddressCfg := 55, [0,55].AlarmCfg := 1, [0,55].AlarmStateCfg := 1, [0,55].OverrideCfg := 1, [0,55].PriorityCfg := 1, [0,55].AlarmONS := 1, [0,56].Tag := 'YA07', [0,56].CurrentValue := 1, [0,56].AlarmCurrentValue := 1, [0,56].AlarmAck := 1, [0,56].Alarm := 1, [0,56].Mimic := 3, [0,56].SoftInput := 1, [0,56].DelayTimer.PRE := 2000, [0,56].DelayTimer.ACC := 2007, [0,56].DelayTimer.EN := 1, [0,56].DelayTimer.DN := 1, [0,56].DelayTimerSP := 2, [0,56].EnableCfg := 1, [0,56].ActiveStateCFg := 1, [0,56].InputAddressCfg := 56, [0,56].AlarmCfg := 1, [0,56].AlarmStateCfg := 1, [0,56].OverrideCfg := 1, [0,56].PriorityCfg := 1, [0,56].AlarmONS := 1, [0,57].Tag := 'YA08', [0,57].DelayTimer.PRE := 5000, [0,57].DelayTimerSP := 5, [0,57].Priority := 1, [0,57].EnableCfg := 1, [0,57].ActiveStateCFg := 1, [0,57].InputAddressCfg := 57, [0,57].AlarmCfg := 1, [0,57].AlarmStateCfg := 1, [0,57].OverrideCfg := 1, [0,57].PriorityCfg := 1, [0,58].Tag := 'YA09', [0,58].CurrentValue := 1, [0,58].AlarmCurrentValue := 1, [0,58].Alarm := 1, [0,58].Mimic := 2, [0,58].SoftInput := 1, [0,58].DelayTimer.PRE := 2000, [0,58].DelayTimer.ACC := 2023, [0,58].DelayTimer.EN := 1, [0,58].DelayTimer.DN := 1,
        [0,58].DelayTimerSP := 2, [0,58].EnableCfg := 1, [0,58].ActiveStateCFg := 1, [0,58].InputAddressCfg := 58, [0,58].AlarmCfg := 1, [0,58].AlarmStateCfg := 1, [0,58].OverrideCfg := 1, [0,58].PriorityCfg := 1, [0,58].AlarmONS := 1, [0,59].Tag := 'YA10', [0,59].CurrentValue := 1, [0,59].Mimic := 1, [0,59].Priority := 1, [0,59].EnableCfg := 1, [0,59].InputAddressCfg := 59, [0,59].AlarmCfg := 1, [0,59].AlarmStateCfg := 1, [0,60].Tag := 'YA11', [0,60].AlarmCurrentValue := 1, [0,60].Override := 1, [0,60].DelayTimer.PRE := 5000, [0,60].DelayTimer.ACC := 2469476, [0,60].DelayTimer.EN := 1, [0,60].DelayTimer.DN := 1, [0,60].DelayTimerSP := 5, [0,60].EnableCfg := 1, [0,60].ActiveStateCFg := 1, [0,60].InputAddressCfg := 60, [0,60].AlarmCfg := 1, [0,60].OverrideCfg := 1, [0,60].PriorityCfg := 1, [0,61].Tag := 'YA12', [0,61].Override := 1, [0,61].DelayTimer.PRE := 2000, [0,61].DelayTimerSP := 2, [0,61].EnableCfg := 1, [0,61].ActiveStateCFg := 1, [0,61].InputAddressCfg := 61, [0,61].AlarmCfg := 1, [0,61].AlarmStateCfg := 1, [0,61].OverrideCfg := 1, [0,61].PriorityCfg := 1, [0,62].Tag := 'UserNCr1', [0,62].CurrentValue := 1, [0,62].Mimic := 1, [0,62].EnableCfg := 1, [0,62].InputAddressCfg := 62, [0,63].Tag := 'UserCr1', [0,63].CurrentValue := 1, [0,63].Mimic := 1, [0,63].Priority := 1, [0,63].EnableCfg := 1, [0,63].InputAddressCfg := 63, [0,64].Tag := 'UserNCr2', [0,64].CurrentValue := 1, [0,64].Mimic := 1, [0,64].EnableCfg := 1, [0,64].InputAddressCfg := 64, [0,65].Tag := 'UserCr2', [0,65].CurrentValue := 1,
        [0,65].Mimic := 1, [0,65].Priority := 1, [0,65].EnableCfg := 1, [0,65].InputAddressCfg := 65, [0,66].Tag := 'LV001_Err', [0,66].DelayTimer.PRE := 2000, [0,66].DelayTimerSP := 2, [0,66].EnableCfg := 1, [0,66].ActiveStateCFg := 1, [0,66].InputAddressCfg := 66, [0,66].AlarmCfg := 1, [0,66].AlarmStateCfg := 1, [0,66].OverrideCfg := 1, [0,66].PriorityCfg := 1, [0,67].Tag := 'LV002_Err', [0,67].DelayTimer.PRE := 2000, [0,67].DelayTimerSP := 2, [0,67].EnableCfg := 1, [0,67].ActiveStateCFg := 1, [0,67].InputAddressCfg := 67, [0,67].AlarmCfg := 1, [0,67].AlarmStateCfg := 1, [0,67].OverrideCfg := 1, [0,67].PriorityCfg := 1, [0,68].CurrentValue := 1, [0,68].AlarmCurrentValue := 1, [0,68].AlarmAck := 1, [0,68].Alarm := 1, [0,68].Mimic := 5, [0,68].SoftInput := 1, [0,68].DelayTimer.PRE := 1000, [0,68].DelayTimer.ACC := 1054, [0,68].DelayTimer.EN := 1, [0,68].DelayTimer.DN := 1, [0,68].DelayTimerSP := 1, [0,68].Priority := 1, [0,68].EnableCfg := 1, [0,68].ActiveStateCFg := 1, [0,68].InputAddressCfg := 68, [0,68].AlarmCfg := 1, [0,68].AlarmStateCfg := 1, [0,68].OverrideCfg := 1, [0,68].AlarmONS := 1, [0,69].CurrentValue := 1, [0,69].AlarmCurrentValue := 1, [0,69].AlarmAck := 1, [0,69].Alarm := 1, [0,69].Mimic := 5, [0,69].SoftInput := 1, [0,69].DelayTimer.PRE := 2000, [0,69].DelayTimer.ACC := 2052, [0,69].DelayTimer.EN := 1, [0,69].DelayTimer.DN := 1, [0,69].DelayTimerSP := 2, [0,69].Priority := 1, [0,69].ActiveStateCFg := 1, [0,69].InputAddressCfg := 69, [0,69].AlarmStateCfg := 1, [0,69].OverrideCfg := 1, [0,69].PriorityCfg := 1,
        [0,69].AlarmONS := 1, [0,70].CurrentValue := 1, [0,70].Mimic := 1, [0,70].DelayTimer.PRE := 2000, [0,70].DelayTimerSP := 2, [0,70].Priority := 1, [0,70].ActiveStateCFg := 1, [0,70].InputAddressCfg := 70, [0,70].AlarmStateCfg := 1, [0,70].OverrideCfg := 1, [0,70].PriorityCfg := 1, [0,71].CurrentValue := 1, [0,71].AlarmCurrentValue := 1, [0,71].AlarmAck := 1, [0,71].Mimic := 5, [0,71].DelayTimer.PRE := 2000, [0,71].DelayTimer.ACC := 2053, [0,71].DelayTimer.EN := 1, [0,71].DelayTimer.DN := 1, [0,71].DelayTimerSP := 2, [0,71].Priority := 1, [0,71].ActiveStateCFg := 1, [0,71].InputAddressCfg := 71, [0,71].AlarmStateCfg := 1, [0,71].OverrideCfg := 1, [0,71].PriorityCfg := 1, [0,71].AlarmONS := 1, [0,72].CurrentValue := 1, [0,72].Mimic := 1, [0,72].DelayTimer.PRE := 2000, [0,72].DelayTimerSP := 2, [0,72].ActiveStateCFg := 1, [0,72].InputAddressCfg := 72, [0,72].AlarmStateCfg := 1, [0,72].OverrideCfg := 1, [0,72].PriorityCfg := 1, [0,73].CurrentValue := 1, [0,73].Mimic := 1, [0,73].DelayTimer.PRE := 2000, [0,73].DelayTimerSP := 2, [0,73].ActiveStateCFg := 1, [0,73].InputAddressCfg := 73, [0,73].AlarmStateCfg := 1, [0,73].OverrideCfg := 1, [0,73].PriorityCfg := 1, [0,74].CurrentValue := 1, [0,74].Mimic := 1, [0,74].DelayTimer.PRE := 2000, [0,74].DelayTimerSP := 2, [0,74].ActiveStateCFg := 1, [0,74].InputAddressCfg := 74, [0,74].AlarmStateCfg := 1, [0,74].OverrideCfg := 1, [0,74].PriorityCfg := 1, [0,75].CurrentValue := 1, [0,75].AlarmCurrentValue := 1, [0,75].AlarmAck := 1, [0,75].Alarm := 1, [0,75].Mimic := 3, [0,75].SoftInput := 1,
        [0,75].DelayTimer.PRE := 2000, [0,75].DelayTimer.ACC := 44, [0,75].DelayTimer.EN := 1, [0,75].DelayTimer.DN := 1, [0,75].DelayTimerSP := 2, [0,75].ActiveStateCFg := 1, [0,75].InputAddressCfg := 75, [0,75].AlarmStateCfg := 1, [0,75].OverrideCfg := 1, [0,75].PriorityCfg := 1, [0,75].AlarmONS := 1, [0,76].CurrentValue := 1, [0,76].Mimic := 1, [0,76].DelayTimer.PRE := 2000, [0,76].DelayTimerSP := 2, [0,76].Priority := 1, [0,76].ActiveStateCFg := 1, [0,76].InputAddressCfg := 76, [0,76].AlarmStateCfg := 1, [0,76].OverrideCfg := 1, [0,76].PriorityCfg := 1, [0,77].CurrentValue := 1, [0,77].Mimic := 1, [0,77].DelayTimer.PRE := 2000, [0,77].DelayTimerSP := 2, [0,77].Priority := 1, [0,77].ActiveStateCFg := 1, [0,77].InputAddressCfg := 77, [0,77].AlarmStateCfg := 1, [0,77].OverrideCfg := 1, [0,77].PriorityCfg := 1, [0,78].CurrentValue := 1, [0,78].AlarmCurrentValue := 1, [0,78].AlarmAck := 1, [0,78].Alarm := 1, [0,78].Mimic := 5, [0,78].SoftInput := 1, [0,78].DelayTimer.PRE := 2000, [0,78].DelayTimer.ACC := 45, [0,78].DelayTimer.EN := 1, [0,78].DelayTimer.DN := 1, [0,78].DelayTimerSP := 2, [0,78].Priority := 1, [0,78].ActiveStateCFg := 1, [0,78].InputAddressCfg := 78, [0,78].AlarmStateCfg := 1, [0,78].OverrideCfg := 1, [0,78].PriorityCfg := 1, [0,78].AlarmONS := 1, [0,79].CurrentValue := 1, [0,79].AlarmCurrentValue := 1, [0,79].Mimic := 1, [0,79].DelayTimer.PRE := 2000, [0,79].DelayTimer.ACC := 44, [0,79].DelayTimer.EN := 1, [0,79].DelayTimer.DN := 1, [0,79].DelayTimerSP := 2, [0,79].Priority := 1, [0,79].ActiveStateCFg := 1, [0,79].InputAddressCfg := 79,
        [0,79].AlarmStateCfg := 1, [0,79].OverrideCfg := 1, [0,79].PriorityCfg := 1, [0,80].CurrentValue := 1, [0,80].AlarmCurrentValue := 1, [0,80].Mimic := 1, [0,80].DelayTimer.PRE := 2000, [0,80].DelayTimer.ACC := 44, [0,80].DelayTimer.EN := 1, [0,80].DelayTimer.DN := 1, [0,80].DelayTimerSP := 2, [0,80].Priority := 1, [0,80].ActiveStateCFg := 1, [0,80].InputAddressCfg := 80, [0,80].AlarmStateCfg := 1, [0,80].OverrideCfg := 1, [0,80].PriorityCfg := 1, [0,81].CurrentValue := 1, [0,81].AlarmCurrentValue := 1, [0,81].Mimic := 1, [0,81].DelayTimer.PRE := 2000, [0,81].DelayTimer.ACC := 44, [0,81].DelayTimer.EN := 1, [0,81].DelayTimer.DN := 1, [0,81].DelayTimerSP := 2, [0,81].ActiveStateCFg := 1, [0,81].InputAddressCfg := 81, [0,81].AlarmStateCfg := 1, [0,81].OverrideCfg := 1, [0,81].PriorityCfg := 1, [0,82].CurrentValue := 1, [0,82].AlarmCurrentValue := 1, [0,82].Mimic := 1, [0,82].DelayTimer.PRE := 2000, [0,82].DelayTimer.ACC := 44, [0,82].DelayTimer.EN := 1, [0,82].DelayTimer.DN := 1, [0,82].DelayTimerSP := 2, [0,82].Priority := 1, [0,82].ActiveStateCFg := 1, [0,82].InputAddressCfg := 82, [0,82].AlarmStateCfg := 1, [0,82].OverrideCfg := 1, [0,82].PriorityCfg := 1, [0,83].CurrentValue := 1, [0,83].AlarmCurrentValue := 1, [0,83].AlarmAck := 1, [0,83].Alarm := 1, [0,83].Mimic := 5, [0,83].SoftInput := 1, [0,83].DelayTimer.PRE := 2000, [0,83].DelayTimer.ACC := 44, [0,83].DelayTimer.EN := 1, [0,83].DelayTimer.DN := 1, [0,83].DelayTimerSP := 2, [0,83].Priority := 1, [0,83].ActiveStateCFg := 1, [0,83].InputAddressCfg := 83, [0,83].AlarmStateCfg := 1, [0,83].OverrideCfg := 1,
        [0,83].PriorityCfg := 1, [0,83].AlarmONS := 1, [0,84].CurrentValue := 1, [0,84].Mimic := 1, [0,84].DelayTimer.PRE := 2000, [0,84].DelayTimerSP := 2, [0,84].Priority := 1, [0,84].ActiveStateCFg := 1, [0,84].InputAddressCfg := 84, [0,84].AlarmStateCfg := 1, [0,84].OverrideCfg := 1, [0,84].PriorityCfg := 1, [0,85].CurrentValue := 1, [0,85].AlarmCurrentValue := 1, [0,85].AlarmAck := 1, [0,85].Alarm := 1, [0,85].Mimic := 3, [0,85].SoftInput := 1, [0,85].DelayTimer.PRE := 2000, [0,85].DelayTimer.ACC := 2021, [0,85].DelayTimer.EN := 1, [0,85].DelayTimer.DN := 1, [0,85].DelayTimerSP := 2, [0,85].ActiveStateCFg := 1, [0,85].InputAddressCfg := 85, [0,85].AlarmStateCfg := 1, [0,85].OverrideCfg := 1, [0,85].PriorityCfg := 1, [0,85].AlarmONS := 1, [0,86].CurrentValue := 1, [0,86].Mimic := 1, [0,86].DelayTimer.PRE := 2000, [0,86].DelayTimerSP := 2, [0,86].ActiveStateCFg := 1, [0,86].InputAddressCfg := 86, [0,86].AlarmStateCfg := 1, [0,86].OverrideCfg := 1, [0,86].PriorityCfg := 1, [0,87].CurrentValue := 1, [0,87].Mimic := 1, [0,87].DelayTimer.PRE := 2000, [0,87].DelayTimerSP := 2, [0,87].ActiveStateCFg := 1, [0,87].InputAddressCfg := 87, [0,87].AlarmStateCfg := 1, [0,87].OverrideCfg := 1, [0,87].PriorityCfg := 1, [0,88].CurrentValue := 1, [0,88].Mimic := 1, [0,88].DelayTimer.PRE := 2000, [0,88].DelayTimerSP := 2, [0,88].ActiveStateCFg := 1, [0,88].InputAddressCfg := 88, [0,88].AlarmStateCfg := 1, [0,88].OverrideCfg := 1, [0,88].PriorityCfg := 1, [0,89].CurrentValue := 1, [0,89].Mimic := 1, [0,89].DelayTimer.PRE := 2000, [0,89].DelayTimerSP := 2,
        [0,89].ActiveStateCFg := 1, [0,89].InputAddressCfg := 89, [0,89].AlarmStateCfg := 1, [0,89].OverrideCfg := 1, [0,89].PriorityCfg := 1, [0,90].Tag := 'PI001_SIG', [0,90].CurrentValue := 1, [0,90].AlarmCurrentValue := 1, [0,90].AlarmAck := 1, [0,90].Alarm := 1, [0,90].Mimic := 5, [0,90].SoftInput := 1, [0,90].DelayTimer.PRE := 2000, [0,90].DelayTimer.ACC := 6308, [0,90].DelayTimer.EN := 1, [0,90].DelayTimer.DN := 1, [0,90].DelayTimerSP := 2, [0,90].Priority := 1, [0,90].EnableCfg := 1, [0,90].ActiveStateCFg := 1, [0,90].InputAddressCfg := 90, [0,90].AlarmCfg := 1, [0,90].AlarmStateCfg := 1, [0,90].OverrideCfg := 1, [0,90].PriorityCfg := 1, [0,90].AlarmONS := 1, [0,91].Tag := 'FI001_SIG', [0,91].DelayTimer.PRE := 2000, [0,91].DelayTimerSP := 2, [0,91].Priority := 1, [0,91].EnableCfg := 1, [0,91].ActiveStateCFg := 1, [0,91].InputAddressCfg := 91, [0,91].AlarmCfg := 1, [0,91].AlarmStateCfg := 1, [0,91].OverrideCfg := 1, [0,91].PriorityCfg := 1, [0,92].Tag := 'PI002_SIG', [0,92].CurrentValue := 1, [0,92].AlarmCurrentValue := 1, [0,92].AlarmAck := 1, [0,92].Alarm := 1, [0,92].Mimic := 5, [0,92].SoftInput := 1, [0,92].DelayTimer.PRE := 2000, [0,92].DelayTimer.EN := 1, [0,92].DelayTimer.DN := 1, [0,92].DelayTimerSP := 2, [0,92].Priority := 1, [0,92].EnableCfg := 1, [0,92].ActiveStateCFg := 1, [0,92].InputAddressCfg := 92, [0,92].AlarmCfg := 1, [0,92].AlarmStateCfg := 1, [0,92].OverrideCfg := 1, [0,92].PriorityCfg := 1, [0,92].AlarmONS := 1, [0,93].Tag := 'FI002_SIG', [0,93].DelayTimer.PRE := 2000, [0,93].DelayTimerSP := 2,
        [0,93].Priority := 1, [0,93].EnableCfg := 1, [0,93].ActiveStateCFg := 1, [0,93].InputAddressCfg := 93, [0,93].AlarmCfg := 1, [0,93].AlarmStateCfg := 1, [0,93].OverrideCfg := 1, [0,93].PriorityCfg := 1, [0,94].Tag := 'PI003_SIG', [0,94].CurrentValue := 1, [0,94].AlarmCurrentValue := 1, [0,94].AlarmAck := 1, [0,94].Alarm := 1, [0,94].Mimic := 3, [0,94].SoftInput := 1, [0,94].DelayTimer.PRE := 2000, [0,94].DelayTimer.ACC := 37, [0,94].DelayTimer.EN := 1, [0,94].DelayTimer.DN := 1, [0,94].DelayTimerSP := 2, [0,94].EnableCfg := 1, [0,94].ActiveStateCFg := 1, [0,94].InputAddressCfg := 94, [0,94].AlarmCfg := 1, [0,94].AlarmStateCfg := 1, [0,94].OverrideCfg := 1, [0,94].PriorityCfg := 1, [0,94].AlarmONS := 1, [0,95].Tag := 'AI102_SIG', [0,95].CurrentValue := 1, [0,95].AlarmCurrentValue := 1, [0,95].AlarmAck := 1, [0,95].Alarm := 1, [0,95].Mimic := 5, [0,95].SoftInput := 1, [0,95].DelayTimer.PRE := 2000, [0,95].DelayTimer.ACC := 2049, [0,95].DelayTimer.EN := 1, [0,95].DelayTimer.DN := 1, [0,95].DelayTimerSP := 2, [0,95].Priority := 1, [0,95].EnableCfg := 1, [0,95].ActiveStateCFg := 1, [0,95].InputAddressCfg := 95, [0,95].AlarmCfg := 1, [0,95].AlarmStateCfg := 1, [0,95].OverrideCfg := 1, [0,95].PriorityCfg := 1, [0,95].AlarmONS := 1, [0,96].Tag := 'AI103_SIG', [0,96].CurrentValue := 1, [0,96].AlarmCurrentValue := 1, [0,96].AlarmAck := 1, [0,96].Alarm := 1, [0,96].Mimic := 5, [0,96].SoftInput := 1, [0,96].DelayTimer.PRE := 2000, [0,96].DelayTimer.ACC := 2049, [0,96].DelayTimer.EN := 1, [0,96].DelayTimer.DN := 1,
        [0,96].DelayTimerSP := 2, [0,96].Priority := 1, [0,96].EnableCfg := 1, [0,96].ActiveStateCFg := 1, [0,96].InputAddressCfg := 96, [0,96].AlarmCfg := 1, [0,96].AlarmStateCfg := 1, [0,96].OverrideCfg := 1, [0,96].PriorityCfg := 1, [0,96].AlarmONS := 1, [0,97].Tag := 'AI201A_SIG', [0,97].CurrentValue := 1, [0,97].AlarmCurrentValue := 1, [0,97].AlarmAck := 1, [0,97].Alarm := 1, [0,97].Mimic := 5, [0,97].SoftInput := 1, [0,97].DelayTimer.PRE := 2000, [0,97].DelayTimer.EN := 1, [0,97].DelayTimer.DN := 1, [0,97].DelayTimerSP := 2, [0,97].Priority := 1, [0,97].EnableCfg := 1, [0,97].ActiveStateCFg := 1, [0,97].InputAddressCfg := 97, [0,97].AlarmCfg := 1, [0,97].AlarmStateCfg := 1, [0,97].OverrideCfg := 1, [0,97].PriorityCfg := 1, [0,97].AlarmONS := 1, [0,98].Tag := 'AI201B_SIG', [0,98].CurrentValue := 1, [0,98].AlarmCurrentValue := 1, [0,98].AlarmAck := 1, [0,98].Alarm := 1, [0,98].Mimic := 5, [0,98].SoftInput := 1, [0,98].DelayTimer.PRE := 2000, [0,98].DelayTimer.EN := 1, [0,98].DelayTimer.DN := 1, [0,98].DelayTimerSP := 2, [0,98].Priority := 1, [0,98].EnableCfg := 1, [0,98].ActiveStateCFg := 1, [0,98].InputAddressCfg := 98, [0,98].AlarmCfg := 1, [0,98].AlarmStateCfg := 1, [0,98].OverrideCfg := 1, [0,98].PriorityCfg := 1, [0,98].AlarmONS := 1, [0,99].Tag := 'TI201_SIG', [0,99].CurrentValue := 1, [0,99].AlarmCurrentValue := 1, [0,99].AlarmAck := 1, [0,99].Alarm := 1, [0,99].Mimic := 3, [0,99].SoftInput := 1, [0,99].DelayTimer.PRE := 2000, [0,99].DelayTimer.EN := 1, [0,99].DelayTimer.DN := 1,
        [0,99].DelayTimerSP := 2, [0,99].EnableCfg := 1, [0,99].ActiveStateCFg := 1, [0,99].InputAddressCfg := 99, [0,99].AlarmCfg := 1, [0,99].AlarmStateCfg := 1, [0,99].OverrideCfg := 1, [0,99].PriorityCfg := 1, [0,99].AlarmONS := 1, [0,100].Tag := 'AI202_SIG', [0,100].CurrentValue := 1, [0,100].AlarmCurrentValue := 1, [0,100].AlarmAck := 1, [0,100].Alarm := 1, [0,100].Mimic := 5, [0,100].SoftInput := 1, [0,100].DelayTimer.PRE := 2000, [0,100].DelayTimer.EN := 1, [0,100].DelayTimer.DN := 1, [0,100].DelayTimerSP := 2, [0,100].Priority := 1, [0,100].EnableCfg := 1, [0,100].ActiveStateCFg := 1, [0,100].InputAddressCfg := 100, [0,100].AlarmCfg := 1, [0,100].AlarmStateCfg := 1, [0,100].OverrideCfg := 1, [0,100].PriorityCfg := 1, [0,100].AlarmONS := 1, [0,101].Tag := 'AI203_SIG', [0,101].CurrentValue := 1, [0,101].AlarmCurrentValue := 1, [0,101].AlarmAck := 1, [0,101].Alarm := 1, [0,101].Mimic := 5, [0,101].SoftInput := 1, [0,101].DelayTimer.PRE := 2000, [0,101].DelayTimer.EN := 1, [0,101].DelayTimer.DN := 1, [0,101].DelayTimerSP := 2, [0,101].Priority := 1, [0,101].EnableCfg := 1, [0,101].ActiveStateCFg := 1, [0,101].InputAddressCfg := 101, [0,101].AlarmCfg := 1, [0,101].AlarmStateCfg := 1, [0,101].OverrideCfg := 1, [0,101].PriorityCfg := 1, [0,101].AlarmONS := 1, [0,102].Tag := 'AI204_SIG', [0,102].CurrentValue := 1, [0,102].AlarmCurrentValue := 1, [0,102].AlarmAck := 1, [0,102].Alarm := 1, [0,102].Mimic := 5, [0,102].SoftInput := 1, [0,102].DelayTimer.PRE := 2000, [0,102].DelayTimer.EN := 1, [0,102].DelayTimer.DN := 1, [0,102].DelayTimerSP := 2,
        [0,102].Priority := 1, [0,102].EnableCfg := 1, [0,102].ActiveStateCFg := 1, [0,102].InputAddressCfg := 102, [0,102].AlarmCfg := 1, [0,102].AlarmStateCfg := 1, [0,102].OverrideCfg := 1, [0,102].PriorityCfg := 1, [0,102].AlarmONS := 1, [0,103].Tag := 'PCV032_SIG', [0,103].CurrentValue := 1, [0,103].AlarmCurrentValue := 1, [0,103].AlarmAck := 1, [0,103].Alarm := 1, [0,103].Mimic := 5, [0,103].SoftInput := 1, [0,103].DelayTimer.PRE := 2000, [0,103].DelayTimer.EN := 1, [0,103].DelayTimer.DN := 1, [0,103].DelayTimerSP := 2, [0,103].Priority := 1, [0,103].EnableCfg := 1, [0,103].ActiveStateCFg := 1, [0,103].InputAddressCfg := 103, [0,103].AlarmCfg := 1, [0,103].AlarmStateCfg := 1, [0,103].OverrideCfg := 1, [0,103].PriorityCfg := 1, [0,103].AlarmONS := 1, [1,0].Tag := 'PSL602', [1,0].CurrentValue := 1, [1,0].Mimic := 1, [1,0].DelayTimer.PRE := 2000, [1,0].DelayTimerSP := 2, [1,0].Priority := 1, [1,0].EnableCfg := 1, [1,0].ActiveStateCFg := 1, [1,0].RealInputCfg := 1, [1,0].AlarmCfg := 1, [1,0].OverrideCfg := 1, [1,0].PriorityCfg := 1, [1,1].Tag := 'XS001', [1,1].CurrentValue := 1, [1,1].Mimic := 1, [1,1].Condition2 := 1, [1,1].DelayTimer.PRE := 1000, [1,1].DelayTimerSP := 1, [1,1].Priority := 1, [1,1].EnableCfg := 1, [1,1].ActiveStateCFg := 1, [1,1].RealInputCfg := 1, [1,1].InputAddressCfg := 1, [1,1].AlarmCfg := 1, [1,1].OverrideCfg := 1, [1,2].Tag := 'XS006', [1,2].DelayTimer.PRE := 1000, [1,2].DelayTimerSP := 1, [1,2].EnableCfg := 1, [1,2].ActiveStateCFg := 1, [1,2].RealInputCfg := 1,
        [1,2].InputAddressCfg := 2, [1,3].Tag := 'ES001', [1,3].CurrentValue := 1, [1,3].Mimic := 1, [1,3].Priority := 1, [1,3].EnableCfg := 1, [1,3].ActiveStateCFg := 1, [1,3].RealInputCfg := 1, [1,3].InputAddressCfg := 3, [1,3].AlarmCfg := 1, [1,4].Tag := 'PSH001', [1,4].CurrentValue := 1, [1,4].Mimic := 1, [1,4].Priority := 1, [1,4].EnableCfg := 1, [1,4].ActiveStateCFg := 1, [1,4].RealInputCfg := 1, [1,4].InputAddressCfg := 4, [1,4].AlarmCfg := 1, [1,4].OverrideCfg := 1, [1,5].Tag := 'PSH401', [1,5].CurrentValue := 1, [1,5].Mimic := 1, [1,5].Priority := 1, [1,5].EnableCfg := 1, [1,5].ActiveStateCFg := 1, [1,5].RealInputCfg := 1, [1,5].InputAddressCfg := 5, [1,5].AlarmCfg := 1, [1,5].OverrideCfg := 1, [1,6].Tag := 'XS002', [1,6].CurrentValue := 1, [1,6].Mimic := 1, [1,6].DelayTimer.PRE := 1000, [1,6].DelayTimerSP := 1, [1,6].EnableCfg := 1, [1,6].ActiveStateCFg := 1, [1,6].RealInputCfg := 1, [1,6].InputAddressCfg := 6, [1,7].Tag := 'XS003', [1,7].CurrentValue := 1, [1,7].Mimic := 1, [1,7].DelayTimer.PRE := 1000, [1,7].DelayTimerSP := 1, [1,7].EnableCfg := 1, [1,7].ActiveStateCFg := 1, [1,7].RealInputCfg := 1, [1,7].InputAddressCfg := 7, [1,8].Tag := 'SIC001DF', [1,8].AlarmCurrentValue := 1, [1,8].AlarmAck := 1, [1,8].Alarm := 1, [1,8].Mimic := 5, [1,8].DelayTimer.PRE := 1000, [1,8].DelayTimer.ACC := 1022, [1,8].DelayTimer.EN := 1, [1,8].DelayTimer.DN := 1, [1,8].DelayTimerSP := 1, [1,8].Priority := 1, [1,8].EnableCfg := 1,
        [1,8].ActiveStateCFg := 1, [1,8].RealInputCfg := 1, [1,8].InputAddressCfg := 8, [1,8].AlarmCfg := 1, [1,8].OverrideCfg := 1, [1,8].PriorityCfg := 1, [1,8].AlarmONS := 1, [1,9].Tag := 'SIC002DF', [1,9].AlarmCurrentValue := 1, [1,9].AlarmAck := 1, [1,9].Alarm := 1, [1,9].Mimic := 5, [1,9].DelayTimer.PRE := 1000, [1,9].DelayTimer.ACC := 1023, [1,9].DelayTimer.EN := 1, [1,9].DelayTimer.DN := 1, [1,9].DelayTimerSP := 1, [1,9].Priority := 1, [1,9].EnableCfg := 1, [1,9].ActiveStateCFg := 1, [1,9].RealInputCfg := 1, [1,9].InputAddressCfg := 9, [1,9].AlarmCfg := 1, [1,9].OverrideCfg := 1, [1,9].PriorityCfg := 1, [1,9].AlarmONS := 1, [1,10].Tag := 'PSL603', [1,10].AlarmCurrentValue := 1, [1,10].AlarmAck := 1, [1,10].Alarm := 1, [1,10].Mimic := 5, [1,10].DelayTimer.PRE := 1000, [1,10].DelayTimer.ACC := 1022, [1,10].DelayTimer.EN := 1, [1,10].DelayTimer.DN := 1, [1,10].DelayTimerSP := 1, [1,10].Priority := 1, [1,10].EnableCfg := 1, [1,10].ActiveStateCFg := 1, [1,10].RealInputCfg := 1, [1,10].InputAddressCfg := 10, [1,10].AlarmCfg := 1, [1,10].OverrideCfg := 1, [1,10].PriorityCfg := 1, [1,10].AlarmONS := 1, [1,11].Tag := 'XS011', [1,11].DelayTimer.PRE := 1000, [1,11].DelayTimerSP := 1, [1,11].ActiveStateCFg := 1, [1,11].RealInputCfg := 1, [1,11].InputAddressCfg := 11, [1,12].Tag := 'XS012', [1,12].DelayTimer.PRE := 1000, [1,12].DelayTimerSP := 1, [1,12].EnableCfg := 1, [1,12].ActiveStateCFg := 1, [1,12].RealInputCfg := 1, [1,12].InputAddressCfg := 12, [1,13].Tag := 'XC102_3DF', [1,13].CurrentValue := 1,
        [1,13].Mimic := 1, [1,13].DelayTimer.PRE := 1000, [1,13].DelayTimerSP := 1, [1,13].Priority := 1, [1,13].EnableCfg := 1, [1,13].ActiveStateCFg := 1, [1,13].RealInputCfg := 1, [1,13].InputAddressCfg := 13, [1,13].AlarmCfg := 1, [1,13].OverrideCfg := 1, [1,13].PriorityCfg := 1, [1,14].Tag := 'SIC003DF', [1,14].AlarmCurrentValue := 1, [1,14].AlarmAck := 1, [1,14].Alarm := 1, [1,14].Mimic := 5, [1,14].DelayTimer.PRE := 1000, [1,14].DelayTimer.ACC := 1022, [1,14].DelayTimer.EN := 1, [1,14].DelayTimer.DN := 1, [1,14].DelayTimerSP := 1, [1,14].Priority := 1, [1,14].EnableCfg := 1, [1,14].ActiveStateCFg := 1, [1,14].RealInputCfg := 1, [1,14].InputAddressCfg := 14, [1,14].AlarmCfg := 1, [1,14].OverrideCfg := 1, [1,14].PriorityCfg := 1, [1,14].AlarmONS := 1, [1,15].Tag := 'SRL001', [1,15].SoftInput := 1, [1,15].DelayTimer.PRE := 2000, [1,15].DelayTimerSP := 2, [1,15].EnableCfg := 1, [1,15].ActiveStateCFg := 1, [1,15].RealInputCfg := 1, [1,15].InputAddressCfg := 15, [1,16].CurrentValue := 1, [1,16].Mimic := 1, [1,16].SoftInput := 1, [1,16].DelayTimer.PRE := 1000, [1,16].DelayTimerSP := 1, [1,16].Priority := 1, [1,16].ActiveStateCFg := 1, [1,16].RealInputCfg := 1, [1,16].InputAddressCfg := 16, [1,16].OverrideCfg := 1, [1,16].PriorityCfg := 1, [1,17].CurrentValue := 1, [1,17].Mimic := 1, [1,17].SoftInput := 1, [1,17].DelayTimer.PRE := 1000, [1,17].DelayTimerSP := 1, [1,17].Priority := 1, [1,17].ActiveStateCFg := 1, [1,17].RealInputCfg := 1, [1,17].InputAddressCfg := 17, [1,17].OverrideCfg := 1, [1,17].PriorityCfg := 1,
        [1,18].CurrentValue := 1, [1,18].Mimic := 1, [1,18].DelayTimer.PRE := 1000, [1,18].DelayTimerSP := 1, [1,18].Priority := 1, [1,18].ActiveStateCFg := 1, [1,18].RealInputCfg := 1, [1,18].InputAddressCfg := 18, [1,18].OverrideCfg := 1, [1,18].PriorityCfg := 1, [1,19].CurrentValue := 1, [1,19].Override := 1, [1,19].Mimic := 1, [1,19].DelayTimer.PRE := 1000, [1,19].DelayTimerSP := 1, [1,19].ActiveStateCFg := 1, [1,19].RealInputCfg := 1, [1,19].InputAddressCfg := 19, [1,19].OverrideCfg := 1, [1,19].PriorityCfg := 1, [1,20].AlarmCurrentValue := 1, [1,20].Override := 1, [1,20].DelayTimer.PRE := 1000, [1,20].DelayTimer.EN := 1, [1,20].DelayTimer.DN := 1, [1,20].DelayTimerSP := 1, [1,20].ActiveStateCFg := 1, [1,20].RealInputCfg := 1, [1,20].InputAddressCfg := 20, [1,20].OverrideCfg := 1, [1,20].PriorityCfg := 1, [1,21].CurrentValue := 1, [1,21].Mimic := 1, [1,21].DelayTimer.PRE := 1000, [1,21].DelayTimerSP := 1, [1,21].Priority := 1, [1,21].ActiveStateCFg := 1, [1,21].RealInputCfg := 1, [1,21].InputAddressCfg := 21, [1,21].OverrideCfg := 1, [1,22].CurrentValue := 1, [1,22].Mimic := 1, [1,22].DelayTimer.PRE := 1000, [1,22].DelayTimerSP := 1, [1,22].Priority := 1, [1,22].ActiveStateCFg := 1, [1,22].RealInputCfg := 1, [1,22].InputAddressCfg := 22, [1,22].OverrideCfg := 1, [1,23].CurrentValue := 1, [1,23].Mimic := 1, [1,23].DelayTimer.PRE := 1000, [1,23].DelayTimerSP := 1, [1,23].Priority := 1, [1,23].ActiveStateCFg := 1, [1,23].RealInputCfg := 1, [1,23].InputAddressCfg := 23, [1,23].OverrideCfg := 1, [1,23].PriorityCfg := 1, [1,24].CurrentValue := 1,
        [1,24].Mimic := 1, [1,24].DelayTimer.PRE := 1000, [1,24].DelayTimerSP := 1, [1,24].Priority := 1, [1,24].ActiveStateCFg := 1, [1,24].RealInputCfg := 1, [1,24].InputAddressCfg := 24, [1,24].OverrideCfg := 1, [1,24].PriorityCfg := 1, [1,25].CurrentValue := 1, [1,25].Mimic := 1, [1,25].DelayTimer.PRE := 20000, [1,25].DelayTimerSP := 2, [1,25].Priority := 1, [1,25].ActiveStateCFg := 1, [1,25].RealInputCfg := 1, [1,25].InputAddressCfg := 25, [1,25].OverrideCfg := 1, [1,25].PriorityCfg := 1, [1,25].Cond1Cfg := 1, [1,26].Override := 1, [1,26].ActiveStateCFg := 1, [1,26].RealInputCfg := 1, [1,26].InputAddressCfg := 26, [1,26].OverrideCfg := 1, [1,26].PriorityCfg := 1, [1,27].Override := 1, [1,27].SoftInput := 1, [1,27].ActiveStateCFg := 1, [1,27].RealInputCfg := 1, [1,27].InputAddressCfg := 27, [1,27].OverrideCfg := 1, [1,27].PriorityCfg := 1, [1,28].Override := 1, [1,28].SoftInput := 1, [1,28].ActiveStateCFg := 1, [1,28].RealInputCfg := 1, [1,28].InputAddressCfg := 28, [1,28].OverrideCfg := 1, [1,28].PriorityCfg := 1, [1,29].Override := 1, [1,29].SoftInput := 1, [1,29].ActiveStateCFg := 1, [1,29].RealInputCfg := 1, [1,29].InputAddressCfg := 29, [1,29].OverrideCfg := 1, [1,29].PriorityCfg := 1, [1,30].Override := 1, [1,30].SoftInput := 1, [1,30].ActiveStateCFg := 1, [1,30].RealInputCfg := 1, [1,30].InputAddressCfg := 30, [1,30].OverrideCfg := 1, [1,30].PriorityCfg := 1, [1,31].Override := 1, [1,31].ActiveStateCFg := 1, [1,31].RealInputCfg := 1, [1,31].InputAddressCfg := 31, [1,31].OverrideCfg := 1, [1,31].PriorityCfg := 1,
        [1,34].Override := 1, [1,34].SoftInput := 1, [1,34].ActiveStateCFg := 1, [1,34].RealInputCfg := 1, [1,34].InputAddressCfg := 34, [1,34].OverrideCfg := 1, [1,34].PriorityCfg := 1, [1,35].Override := 1, [1,35].ActiveStateCFg := 1, [1,35].RealInputCfg := 1, [1,35].InputAddressCfg := 35, [1,35].OverrideCfg := 1, [1,35].PriorityCfg := 1, [1,36].Override := 1, [1,36].SoftInput := 1, [1,36].ActiveStateCFg := 1, [1,36].RealInputCfg := 1, [1,36].InputAddressCfg := 36, [1,36].OverrideCfg := 1, [1,36].PriorityCfg := 1, [1,37].Override := 1, [1,37].ActiveStateCFg := 1, [1,37].RealInputCfg := 1, [1,37].InputAddressCfg := 37, [1,37].OverrideCfg := 1, [1,37].PriorityCfg := 1, [1,38].Override := 1, [1,38].ActiveStateCFg := 1, [1,38].RealInputCfg := 1, [1,38].InputAddressCfg := 38, [1,38].OverrideCfg := 1, [1,38].PriorityCfg := 1, [1,39].Override := 1, [1,39].SoftInput := 1, [1,39].ActiveStateCFg := 1, [1,39].RealInputCfg := 1, [1,39].InputAddressCfg := 39, [1,39].OverrideCfg := 1, [1,39].PriorityCfg := 1, [1,40].Override := 1, [1,40].ActiveStateCFg := 1, [1,40].RealInputCfg := 1, [1,40].InputAddressCfg := 40, [1,40].OverrideCfg := 1, [1,40].PriorityCfg := 1, [1,41].Override := 1, [1,41].SoftInput := 1, [1,41].ActiveStateCFg := 1, [1,41].RealInputCfg := 1, [1,41].InputAddressCfg := 41, [1,41].OverrideCfg := 1, [1,41].PriorityCfg := 1, [1,50].Tag := 'YA01', [1,50].AlarmCurrentValue := 1, [1,50].SoftInput := 1, [1,50].Condition1 := 1, [1,50].DelayTimer.PRE := 60000, [1,50].DelayTimer.ACC := 233, [1,50].DelayTimer.EN := 1, [1,50].DelayTimer.TT := 1,
        [1,50].DelayTimerSP := 60, [1,50].EnableCfg := 1, [1,50].InputAddressCfg := 50, [1,50].AlarmCfg := 1, [1,50].AlarmStateCfg := 1, [1,50].OverrideCfg := 1, [1,50].PriorityCfg := 1, [1,50].Cond1Cfg := 1, [1,51].Tag := 'YA02', [1,51].AlarmCurrentValue := 1, [1,51].SoftInput := 1, [1,51].Condition1 := 1, [1,51].DelayTimer.PRE := 60000, [1,51].DelayTimer.ACC := 31667, [1,51].DelayTimer.EN := 1, [1,51].DelayTimer.TT := 1, [1,51].DelayTimerSP := 60, [1,51].EnableCfg := 1, [1,51].InputAddressCfg := 51, [1,51].AlarmCfg := 1, [1,51].AlarmStateCfg := 1, [1,51].OverrideCfg := 1, [1,51].PriorityCfg := 1, [1,51].Cond1Cfg := 1, [1,52].Tag := 'YA03', [1,52].AlarmCurrentValue := 1, [1,52].SoftInput := 1, [1,52].Condition1 := 1, [1,52].DelayTimer.PRE := 80000, [1,52].DelayTimer.ACC := 31624, [1,52].DelayTimer.EN := 1, [1,52].DelayTimer.TT := 1, [1,52].DelayTimerSP := 80, [1,52].EnableCfg := 1, [1,52].InputAddressCfg := 52, [1,52].AlarmCfg := 1, [1,52].AlarmStateCfg := 1, [1,52].OverrideCfg := 1, [1,52].PriorityCfg := 1, [1,52].Cond1Cfg := 1, [1,53].Tag := 'YA04', [1,53].DelayTimer.PRE := 60000, [1,53].DelayTimerSP := 60, [1,53].EnableCfg := 1, [1,53].ActiveStateCFg := 1, [1,53].InputAddressCfg := 53, [1,53].AlarmCfg := 1, [1,53].AlarmStateCfg := 1, [1,53].OverrideCfg := 1, [1,53].PriorityCfg := 1, [1,54].Tag := 'YA05', [1,54].DelayTimer.PRE := 60000, [1,54].DelayTimerSP := 60, [1,54].EnableCfg := 1, [1,54].ActiveStateCFg := 1, [1,54].InputAddressCfg := 54, [1,54].AlarmCfg := 1, [1,54].AlarmStateCfg := 1, [1,54].OverrideCfg := 1, [1,54].PriorityCfg := 1,
        [1,55].Tag := 'YA06', [1,55].CurrentValue := 1, [1,55].AlarmCurrentValue := 1, [1,55].AlarmAck := 1, [1,55].Alarm := 1, [1,55].Mimic := 5, [1,55].SoftInput := 1, [1,55].DelayTimer.PRE := 5000, [1,55].DelayTimer.ACC := 5004, [1,55].DelayTimer.EN := 1, [1,55].DelayTimer.DN := 1, [1,55].DelayTimerSP := 5, [1,55].Priority := 1, [1,55].EnableCfg := 1, [1,55].ActiveStateCFg := 1, [1,55].InputAddressCfg := 55, [1,55].AlarmCfg := 1, [1,55].AlarmStateCfg := 1, [1,55].OverrideCfg := 1, [1,55].PriorityCfg := 1, [1,55].AlarmONS := 1, [1,56].Tag := 'YA07', [1,56].DelayTimer.PRE := 2000, [1,56].DelayTimerSP := 2, [1,56].EnableCfg := 1, [1,56].ActiveStateCFg := 1, [1,56].InputAddressCfg := 56, [1,56].AlarmCfg := 1, [1,56].AlarmStateCfg := 1, [1,56].OverrideCfg := 1, [1,56].PriorityCfg := 1, [1,57].Tag := 'YA08', [1,57].DelayTimer.PRE := 5000, [1,57].DelayTimerSP := 5, [1,57].Priority := 1, [1,57].EnableCfg := 1, [1,57].ActiveStateCFg := 1, [1,57].InputAddressCfg := 57, [1,57].AlarmCfg := 1, [1,57].AlarmStateCfg := 1, [1,57].OverrideCfg := 1, [1,57].PriorityCfg := 1, [1,58].Tag := 'YA09', [1,58].DelayTimer.PRE := 2000, [1,58].DelayTimerSP := 2, [1,58].EnableCfg := 1, [1,58].ActiveStateCFg := 1, [1,58].InputAddressCfg := 58, [1,58].AlarmCfg := 1, [1,58].AlarmStateCfg := 1, [1,58].OverrideCfg := 1, [1,58].PriorityCfg := 1, [1,59].Tag := 'YA10', [1,59].CurrentValue := 1, [1,59].Mimic := 1, [1,59].Priority := 1, [1,59].EnableCfg := 1, [1,59].InputAddressCfg := 59, [1,59].AlarmCfg := 1, [1,59].AlarmStateCfg := 1,
        [1,60].Tag := 'YA11', [1,60].Override := 1, [1,60].DelayTimer.PRE := 5000, [1,60].DelayTimerSP := 5, [1,60].EnableCfg := 1, [1,60].ActiveStateCFg := 1, [1,60].InputAddressCfg := 60, [1,60].AlarmCfg := 1, [1,60].AlarmStateCfg := 1, [1,60].OverrideCfg := 1, [1,60].PriorityCfg := 1, [1,61].Tag := 'YA12', [1,61].EnableCfg := 1, [1,61].ActiveStateCFg := 1, [1,61].InputAddressCfg := 61, [1,61].AlarmCfg := 1, [1,61].AlarmStateCfg := 1, [1,61].OverrideCfg := 1, [1,61].PriorityCfg := 1, [1,62].Tag := 'YA13', [1,62].CurrentValue := 1, [1,62].AlarmCurrentValue := 1, [1,62].AlarmAck := 1, [1,62].Alarm := 1, [1,62].Mimic := 3, [1,62].SoftInput := 1, [1,62].DelayTimer.PRE := 2000, [1,62].DelayTimer.ACC := 2005, [1,62].DelayTimer.EN := 1, [1,62].DelayTimer.DN := 1, [1,62].DelayTimerSP := 2, [1,62].EnableCfg := 1, [1,62].ActiveStateCFg := 1, [1,62].InputAddressCfg := 62, [1,62].AlarmCfg := 1, [1,62].AlarmStateCfg := 1, [1,62].OverrideCfg := 1, [1,62].PriorityCfg := 1, [1,62].AlarmONS := 1, [1,63].Tag := 'YA14', [1,63].CurrentValue := 1, [1,63].Mimic := 1, [1,63].DelayTimer.PRE := 60000, [1,63].DelayTimerSP := 60, [1,63].EnableCfg := 1, [1,63].InputAddressCfg := 63, [1,63].AlarmCfg := 1, [1,63].AlarmStateCfg := 1, [1,64].Tag := 'UserNCr1', [1,64].CurrentValue := 1, [1,64].Mimic := 1, [1,64].EnableCfg := 1, [1,64].InputAddressCfg := 64, [1,65].Tag := 'UserCr1', [1,65].CurrentValue := 1, [1,65].Mimic := 1, [1,65].Priority := 1, [1,65].EnableCfg := 1, [1,65].InputAddressCfg := 65, [1,66].Tag := 'UserNCr2',
        [1,66].CurrentValue := 1, [1,66].Mimic := 1, [1,66].DelayTimer.PRE := 2000, [1,66].DelayTimerSP := 2, [1,66].EnableCfg := 1, [1,66].InputAddressCfg := 66, [1,67].Tag := 'UserCr2', [1,67].CurrentValue := 1, [1,67].Mimic := 1, [1,67].DelayTimer.PRE := 2000, [1,67].DelayTimerSP := 2, [1,67].Priority := 1, [1,67].EnableCfg := 1, [1,67].InputAddressCfg := 67, [1,68].Tag := 'ZSDF', [1,68].CurrentValue := 1, [1,68].AlarmCurrentValue := 1, [1,68].AlarmAck := 1, [1,68].Alarm := 1, [1,68].Mimic := 5, [1,68].SoftInput := 1, [1,68].DelayTimer.PRE := 1000, [1,68].DelayTimer.ACC := 1028, [1,68].DelayTimer.EN := 1, [1,68].DelayTimer.DN := 1, [1,68].DelayTimerSP := 1, [1,68].Priority := 1, [1,68].EnableCfg := 1, [1,68].ActiveStateCFg := 1, [1,68].InputAddressCfg := 68, [1,68].AlarmCfg := 1, [1,68].AlarmStateCfg := 1, [1,68].OverrideCfg := 1, [1,68].PriorityCfg := 1, [1,68].AlarmONS := 1, [1,69].Tag := 'YA15', [1,69].CurrentValue := 1, [1,69].AlarmCurrentValue := 1, [1,69].AlarmAck := 1, [1,69].Alarm := 1, [1,69].Mimic := 5, [1,69].SoftInput := 1, [1,69].DelayTimer.PRE := 5000, [1,69].DelayTimer.EN := 1, [1,69].DelayTimer.DN := 1, [1,69].DelayTimerSP := 5, [1,69].Priority := 1, [1,69].EnableCfg := 1, [1,69].ActiveStateCFg := 1, [1,69].InputAddressCfg := 69, [1,69].AlarmCfg := 1, [1,69].AlarmStateCfg := 1, [1,69].OverrideCfg := 1, [1,69].PriorityCfg := 1, [1,69].AlarmONS := 1, [1,70].Tag := 'YA16', [1,70].DelayTimer.PRE := 2000, [1,70].DelayTimerSP := 2, [1,70].EnableCfg := 1, [1,70].ActiveStateCFg := 1,
        [1,70].InputAddressCfg := 70, [1,70].AlarmCfg := 1, [1,70].AlarmStateCfg := 1, [1,70].OverrideCfg := 1, [1,70].PriorityCfg := 1, [1,71].Tag := 'YA17', [1,71].DelayTimer.PRE := 5000, [1,71].DelayTimerSP := 5, [1,71].Priority := 1, [1,71].EnableCfg := 1, [1,71].ActiveStateCFg := 1, [1,71].InputAddressCfg := 71, [1,71].AlarmCfg := 1, [1,71].AlarmStateCfg := 1, [1,71].OverrideCfg := 1, [1,71].PriorityCfg := 1, [1,72].Tag := 'YA18', [1,72].DelayTimer.PRE := 2000, [1,72].DelayTimerSP := 2, [1,72].EnableCfg := 1, [1,72].ActiveStateCFg := 1, [1,72].InputAddressCfg := 72, [1,72].AlarmCfg := 1, [1,72].AlarmStateCfg := 1, [1,72].OverrideCfg := 1, [1,72].PriorityCfg := 1, [1,73].Tag := 'YA19', [1,73].DelayTimer.PRE := 5000, [1,73].DelayTimerSP := 5, [1,73].Priority := 1, [1,73].EnableCfg := 1, [1,73].ActiveStateCFg := 1, [1,73].InputAddressCfg := 73, [1,73].AlarmCfg := 1, [1,73].AlarmStateCfg := 1, [1,73].OverrideCfg := 1, [1,73].PriorityCfg := 1, [1,74].Tag := 'YA20', [1,74].DelayTimer.PRE := 2000, [1,74].DelayTimerSP := 2, [1,74].EnableCfg := 1, [1,74].ActiveStateCFg := 1, [1,74].InputAddressCfg := 74, [1,74].AlarmCfg := 1, [1,74].AlarmStateCfg := 1, [1,74].OverrideCfg := 1, [1,74].PriorityCfg := 1, [1,75].Tag := 'YA21', [1,75].DelayTimer.PRE := 5000, [1,75].DelayTimerSP := 5, [1,75].Priority := 1, [1,75].EnableCfg := 1, [1,75].ActiveStateCFg := 1, [1,75].InputAddressCfg := 75, [1,75].AlarmCfg := 1, [1,75].AlarmStateCfg := 1, [1,75].OverrideCfg := 1, [1,75].PriorityCfg := 1, [1,76].Tag := 'YA41', [1,76].DelayTimer.PRE := 5000,
        [1,76].DelayTimerSP := 5, [1,76].Priority := 1, [1,76].EnableCfg := 1, [1,76].ActiveStateCFg := 1, [1,76].InputAddressCfg := 76, [1,76].AlarmCfg := 1, [1,76].AlarmStateCfg := 1, [1,76].OverrideCfg := 1, [1,76].PriorityCfg := 1, [1,77].EnableCfg := 1, [1,77].ActiveStateCFg := 1, [1,77].InputAddressCfg := 77, [1,77].AlarmCfg := 1, [1,77].AlarmStateCfg := 1, [1,77].OverrideCfg := 1, [1,78].CurrentValue := 1, [1,78].AlarmCurrentValue := 1, [1,78].AlarmAck := 1, [1,78].Alarm := 1, [1,78].Mimic := 5, [1,78].SoftInput := 1, [1,78].DelayTimer.PRE := 2000, [1,78].DelayTimer.ACC := 45, [1,78].DelayTimer.EN := 1, [1,78].DelayTimer.DN := 1, [1,78].DelayTimerSP := 2, [1,78].Priority := 1, [1,78].ActiveStateCFg := 1, [1,78].InputAddressCfg := 78, [1,78].AlarmStateCfg := 1, [1,78].OverrideCfg := 1, [1,78].PriorityCfg := 1, [1,78].AlarmONS := 1, [1,79].CurrentValue := 1, [1,79].AlarmCurrentValue := 1, [1,79].Mimic := 1, [1,79].DelayTimer.PRE := 2000, [1,79].DelayTimer.ACC := 44, [1,79].DelayTimer.EN := 1, [1,79].DelayTimer.DN := 1, [1,79].DelayTimerSP := 2, [1,79].Priority := 1, [1,79].ActiveStateCFg := 1, [1,79].InputAddressCfg := 79, [1,79].AlarmStateCfg := 1, [1,79].OverrideCfg := 1, [1,79].PriorityCfg := 1, [1,80].CurrentValue := 1, [1,80].AlarmCurrentValue := 1, [1,80].Mimic := 1, [1,80].DelayTimer.PRE := 2000, [1,80].DelayTimer.ACC := 44, [1,80].DelayTimer.EN := 1, [1,80].DelayTimer.DN := 1, [1,80].DelayTimerSP := 2, [1,80].Priority := 1, [1,80].ActiveStateCFg := 1, [1,80].InputAddressCfg := 80, [1,80].AlarmStateCfg := 1, [1,80].OverrideCfg := 1,
        [1,80].PriorityCfg := 1, [1,81].CurrentValue := 1, [1,81].AlarmCurrentValue := 1, [1,81].Mimic := 1, [1,81].DelayTimer.PRE := 2000, [1,81].DelayTimer.ACC := 44, [1,81].DelayTimer.EN := 1, [1,81].DelayTimer.DN := 1, [1,81].DelayTimerSP := 2, [1,81].ActiveStateCFg := 1, [1,81].InputAddressCfg := 81, [1,81].AlarmStateCfg := 1, [1,81].OverrideCfg := 1, [1,81].PriorityCfg := 1, [1,82].CurrentValue := 1, [1,82].AlarmCurrentValue := 1, [1,82].Mimic := 1, [1,82].DelayTimer.PRE := 2000, [1,82].DelayTimer.ACC := 44, [1,82].DelayTimer.EN := 1, [1,82].DelayTimer.DN := 1, [1,82].DelayTimerSP := 2, [1,82].Priority := 1, [1,82].ActiveStateCFg := 1, [1,82].InputAddressCfg := 82, [1,82].AlarmStateCfg := 1, [1,82].OverrideCfg := 1, [1,82].PriorityCfg := 1, [1,83].CurrentValue := 1, [1,83].AlarmCurrentValue := 1, [1,83].AlarmAck := 1, [1,83].Alarm := 1, [1,83].Mimic := 5, [1,83].SoftInput := 1, [1,83].DelayTimer.PRE := 2000, [1,83].DelayTimer.ACC := 44, [1,83].DelayTimer.EN := 1, [1,83].DelayTimer.DN := 1, [1,83].DelayTimerSP := 2, [1,83].Priority := 1, [1,83].ActiveStateCFg := 1, [1,83].InputAddressCfg := 83, [1,83].AlarmStateCfg := 1, [1,83].OverrideCfg := 1, [1,83].PriorityCfg := 1, [1,83].AlarmONS := 1, [1,84].CurrentValue := 1, [1,84].Mimic := 1, [1,84].DelayTimer.PRE := 2000, [1,84].DelayTimerSP := 2, [1,84].Priority := 1, [1,84].ActiveStateCFg := 1, [1,84].InputAddressCfg := 84, [1,84].AlarmStateCfg := 1, [1,84].OverrideCfg := 1, [1,84].PriorityCfg := 1, [1,85].CurrentValue := 1, [1,85].AlarmCurrentValue := 1, [1,85].AlarmAck := 1, [1,85].Alarm := 1,
        [1,85].Mimic := 3, [1,85].SoftInput := 1, [1,85].DelayTimer.PRE := 2000, [1,85].DelayTimer.ACC := 2021, [1,85].DelayTimer.EN := 1, [1,85].DelayTimer.DN := 1, [1,85].DelayTimerSP := 2, [1,85].ActiveStateCFg := 1, [1,85].InputAddressCfg := 85, [1,85].AlarmStateCfg := 1, [1,85].OverrideCfg := 1, [1,85].PriorityCfg := 1, [1,85].AlarmONS := 1, [1,86].CurrentValue := 1, [1,86].Mimic := 1, [1,86].DelayTimer.PRE := 2000, [1,86].DelayTimerSP := 2, [1,86].ActiveStateCFg := 1, [1,86].InputAddressCfg := 86, [1,86].AlarmStateCfg := 1, [1,86].OverrideCfg := 1, [1,86].PriorityCfg := 1, [1,87].CurrentValue := 1, [1,87].Mimic := 1, [1,87].DelayTimer.PRE := 2000, [1,87].DelayTimerSP := 2, [1,87].ActiveStateCFg := 1, [1,87].InputAddressCfg := 87, [1,87].AlarmStateCfg := 1, [1,87].OverrideCfg := 1, [1,87].PriorityCfg := 1, [1,88].CurrentValue := 1, [1,88].Mimic := 1, [1,88].DelayTimer.PRE := 2000, [1,88].DelayTimerSP := 2, [1,88].ActiveStateCFg := 1, [1,88].InputAddressCfg := 88, [1,88].AlarmStateCfg := 1, [1,88].OverrideCfg := 1, [1,88].PriorityCfg := 1, [1,89].CurrentValue := 1, [1,89].Mimic := 1, [1,89].DelayTimer.PRE := 2000, [1,89].DelayTimerSP := 2, [1,89].ActiveStateCFg := 1, [1,89].InputAddressCfg := 89, [1,89].AlarmStateCfg := 1, [1,89].OverrideCfg := 1, [1,89].PriorityCfg := 1, [1,90].Tag := 'AI101_SIG', [1,90].DelayTimer.PRE := 2000, [1,90].DelayTimerSP := 2, [1,90].EnableCfg := 1, [1,90].ActiveStateCFg := 1, [1,90].InputAddressCfg := 90, [1,90].AlarmCfg := 1, [1,90].AlarmStateCfg := 1, [1,90].OverrideCfg := 1, [1,90].PriorityCfg := 1, [1,91].Tag := 'AI102_SIG',
        [1,91].DelayTimer.PRE := 10000, [1,91].DelayTimerSP := 10, [1,91].EnableCfg := 1, [1,91].ActiveStateCFg := 1, [1,91].InputAddressCfg := 91, [1,91].AlarmCfg := 1, [1,91].AlarmStateCfg := 1, [1,91].OverrideCfg := 1, [1,91].PriorityCfg := 1, [1,92].Tag := 'AI103_SIG', [1,92].DelayTimer.PRE := 10000, [1,92].DelayTimerSP := 10, [1,92].EnableCfg := 1, [1,92].ActiveStateCFg := 1, [1,92].InputAddressCfg := 92, [1,92].AlarmCfg := 1, [1,92].AlarmStateCfg := 1, [1,92].OverrideCfg := 1, [1,92].PriorityCfg := 1, [1,93].Tag := 'FI101_SIG', [1,93].DelayTimer.PRE := 10000, [1,93].DelayTimerSP := 10, [1,93].EnableCfg := 1, [1,93].ActiveStateCFg := 1, [1,93].InputAddressCfg := 93, [1,93].AlarmCfg := 1, [1,93].AlarmStateCfg := 1, [1,93].OverrideCfg := 1, [1,93].PriorityCfg := 1, [1,94].Tag := 'WI001_SIG', [1,94].DelayTimer.PRE := 10000, [1,94].DelayTimerSP := 10, [1,94].EnableCfg := 1, [1,94].ActiveStateCFg := 1, [1,94].InputAddressCfg := 94, [1,94].AlarmCfg := 1, [1,94].AlarmStateCfg := 1, [1,94].OverrideCfg := 1, [1,94].PriorityCfg := 1, [1,95].Tag := 'WI101_SIG', [1,95].DelayTimer.PRE := 10000, [1,95].DelayTimerSP := 10, [1,95].EnableCfg := 1, [1,95].ActiveStateCFg := 1, [1,95].InputAddressCfg := 95, [1,95].AlarmCfg := 1, [1,95].AlarmStateCfg := 1, [1,95].OverrideCfg := 1, [1,95].PriorityCfg := 1, [1,96].Tag := 'WI102_SIG', [1,96].CurrentValue := 1, [1,96].AlarmCurrentValue := 1, [1,96].AlarmAck := 1, [1,96].Mimic := 5, [1,96].SoftInput := 1, [1,96].DelayTimer.PRE := 2000, [1,96].DelayTimer.ACC := 2021, [1,96].DelayTimer.EN := 1, [1,96].DelayTimer.DN := 1, [1,96].DelayTimerSP := 2,
        [1,96].ActiveStateCFg := 1, [1,96].InputAddressCfg := 96, [1,96].AlarmStateCfg := 1, [1,96].OverrideCfg := 1, [1,96].PriorityCfg := 1, [1,96].AlarmONS := 1, [1,97].Tag := 'PI001_SIG', [1,97].DelayTimer.PRE := 10000, [1,97].DelayTimerSP := 10, [1,97].EnableCfg := 1, [1,97].ActiveStateCFg := 1, [1,97].InputAddressCfg := 97, [1,97].AlarmCfg := 1, [1,97].AlarmStateCfg := 1, [1,97].OverrideCfg := 1, [1,97].PriorityCfg := 1, [1,98].Tag := 'PI002_SIG', [1,98].DelayTimer.PRE := 10000, [1,98].DelayTimerSP := 10, [1,98].EnableCfg := 1, [1,98].ActiveStateCFg := 1, [1,98].InputAddressCfg := 98, [1,98].AlarmCfg := 1, [1,98].AlarmStateCfg := 1, [1,98].OverrideCfg := 1, [1,98].PriorityCfg := 1, [1,99].Tag := 'PI101_SIG', [1,99].DelayTimer.PRE := 10000, [1,99].DelayTimerSP := 10, [1,99].EnableCfg := 1, [1,99].ActiveStateCFg := 1, [1,99].InputAddressCfg := 99, [1,99].AlarmCfg := 1, [1,99].AlarmStateCfg := 1, [1,99].OverrideCfg := 1, [1,99].PriorityCfg := 1, [1,100].Tag := 'PI401_SIG', [1,100].DelayTimer.PRE := 10000, [1,100].DelayTimerSP := 10, [1,100].EnableCfg := 1, [1,100].ActiveStateCFg := 1, [1,100].InputAddressCfg := 100, [1,100].AlarmCfg := 1, [1,100].AlarmStateCfg := 1, [1,100].OverrideCfg := 1, [1,100].PriorityCfg := 1, [1,101].Tag := 'TI001_SIG', [1,101].DelayTimer.PRE := 10000, [1,101].DelayTimerSP := 10, [1,101].EnableCfg := 1, [1,101].ActiveStateCFg := 1, [1,101].InputAddressCfg := 101, [1,101].AlarmCfg := 1, [1,101].AlarmStateCfg := 1, [1,101].OverrideCfg := 1, [1,101].PriorityCfg := 1, [1,102].Tag := 'PCV001_SIG', [1,102].DelayTimer.PRE := 10000, [1,102].DelayTimerSP := 10, [1,102].EnableCfg := 1,
        [1,102].ActiveStateCFg := 1, [1,102].InputAddressCfg := 102, [1,102].AlarmCfg := 1, [1,102].AlarmStateCfg := 1, [1,102].OverrideCfg := 1, [1,102].PriorityCfg := 1, [1,103].Tag := 'PCV101_SIG', [1,103].DelayTimer.PRE := 10000, [1,103].DelayTimerSP := 10, [1,103].EnableCfg := 1, [1,103].ActiveStateCFg := 1, [1,103].InputAddressCfg := 103, [1,103].AlarmCfg := 1, [1,103].AlarmStateCfg := 1, [1,103].OverrideCfg := 1, [1,103].PriorityCfg := 1, [1,104].Tag := 'MIX001_SIG', [1,104].DelayTimer.PRE := 10000, [1,104].DelayTimerSP := 10, [1,104].EnableCfg := 1, [1,104].ActiveStateCFg := 1, [1,104].InputAddressCfg := 104, [1,104].AlarmCfg := 1, [1,104].AlarmStateCfg := 1, [1,104].OverrideCfg := 1, [1,104].PriorityCfg := 1, [1,105].Tag := 'AI104_SIG', [1,105].CurrentValue := 1, [1,105].AlarmCurrentValue := 1, [1,105].Mimic := 4, [1,105].SoftInput := 1, [1,105].DelayTimer.PRE := 2000, [1,105].DelayTimer.ACC := 40, [1,105].DelayTimer.EN := 1, [1,105].DelayTimer.DN := 1, [1,105].DelayTimerSP := 10, [1,105].ActiveStateCFg := 1, [1,105].InputAddressCfg := 105, [1,105].AlarmStateCfg := 1, [1,105].OverrideCfg := 1, [1,105].PriorityCfg := 1, [1,105].AlarmONS := 1, [1,106].Tag := 'FI003_SIG', [1,106].SoftInput := 1, [1,106].DelayTimerSP := 10, [1,106].ActiveStateCFg := 1, [1,106].InputAddressCfg := 106, [1,106].AlarmStateCfg := 1, [1,106].OverrideCfg := 1, [1,106].PriorityCfg := 1, [2,0].Tag := 'PSL602', [2,0].CurrentValue := 1, [2,0].Mimic := 1, [2,0].DelayTimer.PRE := 2000, [2,0].DelayTimerSP := 2, [2,0].Priority := 1, [2,0].EnableCfg := 1, [2,0].ActiveStateCFg := 1, [2,0].RealInputCfg := 1, [2,0].AlarmCfg := 1,
        [2,0].OverrideCfg := 1, [2,0].PriorityCfg := 1, [2,1].Tag := 'XS001', [2,1].CurrentValue := 1, [2,1].Mimic := 1, [2,1].Condition2 := 1, [2,1].DelayTimer.PRE := 1000, [2,1].DelayTimerSP := 1, [2,1].Priority := 1, [2,1].EnableCfg := 1, [2,1].ActiveStateCFg := 1, [2,1].RealInputCfg := 1, [2,1].InputAddressCfg := 1, [2,1].AlarmCfg := 1, [2,1].OverrideCfg := 1, [2,2].Tag := 'XS006', [2,2].DelayTimer.PRE := 1000, [2,2].DelayTimerSP := 1, [2,2].EnableCfg := 1, [2,2].ActiveStateCFg := 1, [2,2].RealInputCfg := 1, [2,2].InputAddressCfg := 2, [2,3].Tag := 'ES001', [2,3].CurrentValue := 1, [2,3].Mimic := 1, [2,3].Priority := 1, [2,3].EnableCfg := 1, [2,3].ActiveStateCFg := 1, [2,3].RealInputCfg := 1, [2,3].InputAddressCfg := 3, [2,3].AlarmCfg := 1, [2,4].Tag := 'PSH001', [2,4].AlarmCurrentValue := 1, [2,4].Alarm := 1, [2,4].Mimic := 4, [2,4].DelayTimer.ACC := 52, [2,4].DelayTimer.EN := 1, [2,4].DelayTimer.DN := 1, [2,4].Priority := 1, [2,4].EnableCfg := 1, [2,4].ActiveStateCFg := 1, [2,4].RealInputCfg := 1, [2,4].InputAddressCfg := 4, [2,4].AlarmCfg := 1, [2,4].OverrideCfg := 1, [2,4].AlarmONS := 1, [2,5].Tag := 'PSH401', [2,5].AlarmCurrentValue := 1, [2,5].Alarm := 1, [2,5].Mimic := 4, [2,5].DelayTimer.ACC := 52, [2,5].DelayTimer.EN := 1, [2,5].DelayTimer.DN := 1, [2,5].Priority := 1, [2,5].EnableCfg := 1, [2,5].ActiveStateCFg := 1, [2,5].RealInputCfg := 1, [2,5].InputAddressCfg := 5, [2,5].AlarmCfg := 1, [2,5].OverrideCfg := 1,
        [2,5].AlarmONS := 1, [2,6].Tag := 'XS002', [2,6].DelayTimer.PRE := 1000, [2,6].DelayTimerSP := 1, [2,6].EnableCfg := 1, [2,6].ActiveStateCFg := 1, [2,6].RealInputCfg := 1, [2,6].InputAddressCfg := 6, [2,7].Tag := 'XS003', [2,7].DelayTimer.PRE := 1000, [2,7].DelayTimerSP := 1, [2,7].EnableCfg := 1, [2,7].ActiveStateCFg := 1, [2,7].RealInputCfg := 1, [2,7].InputAddressCfg := 7, [2,8].Tag := 'SIC001DF', [2,8].AlarmCurrentValue := 1, [2,8].AlarmAck := 1, [2,8].Alarm := 1, [2,8].Mimic := 5, [2,8].DelayTimer.PRE := 1000, [2,8].DelayTimer.ACC := 1039, [2,8].DelayTimer.EN := 1, [2,8].DelayTimer.DN := 1, [2,8].DelayTimerSP := 1, [2,8].Priority := 1, [2,8].EnableCfg := 1, [2,8].ActiveStateCFg := 1, [2,8].RealInputCfg := 1, [2,8].InputAddressCfg := 8, [2,8].AlarmCfg := 1, [2,8].OverrideCfg := 1, [2,8].PriorityCfg := 1, [2,8].AlarmONS := 1, [2,9].Tag := 'SIC002DF', [2,9].AlarmCurrentValue := 1, [2,9].AlarmAck := 1, [2,9].Alarm := 1, [2,9].Mimic := 5, [2,9].DelayTimer.PRE := 1000, [2,9].DelayTimer.ACC := 1038, [2,9].DelayTimer.EN := 1, [2,9].DelayTimer.DN := 1, [2,9].DelayTimerSP := 1, [2,9].Priority := 1, [2,9].EnableCfg := 1, [2,9].ActiveStateCFg := 1, [2,9].RealInputCfg := 1, [2,9].InputAddressCfg := 9, [2,9].AlarmCfg := 1, [2,9].OverrideCfg := 1, [2,9].PriorityCfg := 1, [2,9].AlarmONS := 1, [2,10].Tag := 'PSL603', [2,10].AlarmCurrentValue := 1, [2,10].AlarmAck := 1, [2,10].Alarm := 1, [2,10].Mimic := 5, [2,10].DelayTimer.PRE := 1000, [2,10].DelayTimer.ACC := 1038,
        [2,10].DelayTimer.EN := 1, [2,10].DelayTimer.DN := 1, [2,10].DelayTimerSP := 1, [2,10].Priority := 1, [2,10].EnableCfg := 1, [2,10].ActiveStateCFg := 1, [2,10].RealInputCfg := 1, [2,10].InputAddressCfg := 10, [2,10].AlarmCfg := 1, [2,10].OverrideCfg := 1, [2,10].PriorityCfg := 1, [2,10].AlarmONS := 1, [2,11].Tag := 'XS011', [2,11].DelayTimer.PRE := 1000, [2,11].DelayTimerSP := 1, [2,11].EnableCfg := 1, [2,11].ActiveStateCFg := 1, [2,11].RealInputCfg := 1, [2,11].InputAddressCfg := 11, [2,12].Tag := 'XS012', [2,12].DelayTimer.PRE := 1000, [2,12].DelayTimerSP := 1, [2,12].EnableCfg := 1, [2,12].ActiveStateCFg := 1, [2,12].RealInputCfg := 1, [2,12].InputAddressCfg := 12, [2,13].Tag := 'XC102_3DF', [2,13].CurrentValue := 1, [2,13].Mimic := 1, [2,13].DelayTimer.PRE := 20000, [2,13].DelayTimerSP := 1, [2,13].Priority := 1, [2,13].ActiveStateCFg := 1, [2,13].RealInputCfg := 1, [2,13].InputAddressCfg := 13, [2,13].OverrideCfg := 1, [2,13].PriorityCfg := 1, [2,14].Tag := 'SIC003DF', [2,14].AlarmCurrentValue := 1, [2,14].AlarmAck := 1, [2,14].Alarm := 1, [2,14].Mimic := 5, [2,14].DelayTimer.PRE := 1000, [2,14].DelayTimer.ACC := 1039, [2,14].DelayTimer.EN := 1, [2,14].DelayTimer.DN := 1, [2,14].DelayTimerSP := 1, [2,14].Priority := 1, [2,14].EnableCfg := 1, [2,14].ActiveStateCFg := 1, [2,14].RealInputCfg := 1, [2,14].InputAddressCfg := 14, [2,14].AlarmCfg := 1, [2,14].OverrideCfg := 1, [2,14].PriorityCfg := 1, [2,14].AlarmONS := 1, [2,15].Tag := 'SRL001', [2,15].SoftInput := 1, [2,15].DelayTimer.PRE := 2000, [2,15].DelayTimerSP := 2,
        [2,15].EnableCfg := 1, [2,15].ActiveStateCFg := 1, [2,15].RealInputCfg := 1, [2,15].InputAddressCfg := 15, [2,16].AlarmCurrentValue := 1, [2,16].Override := 1, [2,16].SoftInput := 1, [2,16].DelayTimer.PRE := 1000, [2,16].DelayTimer.ACC := 1018, [2,16].DelayTimer.EN := 1, [2,16].DelayTimer.DN := 1, [2,16].DelayTimerSP := 1, [2,16].Priority := 1, [2,16].ActiveStateCFg := 1, [2,16].RealInputCfg := 1, [2,16].InputAddressCfg := 16, [2,16].OverrideCfg := 1, [2,16].PriorityCfg := 1, [2,17].AlarmCurrentValue := 1, [2,17].Override := 1, [2,17].SoftInput := 1, [2,17].DelayTimer.PRE := 1000, [2,17].DelayTimer.ACC := 1018, [2,17].DelayTimer.EN := 1, [2,17].DelayTimer.DN := 1, [2,17].DelayTimerSP := 1, [2,17].Priority := 1, [2,17].ActiveStateCFg := 1, [2,17].RealInputCfg := 1, [2,17].InputAddressCfg := 17, [2,17].OverrideCfg := 1, [2,17].PriorityCfg := 1, [2,18].AlarmCurrentValue := 1, [2,18].Override := 1, [2,18].DelayTimer.PRE := 1000, [2,18].DelayTimer.ACC := 1018, [2,18].DelayTimer.EN := 1, [2,18].DelayTimer.DN := 1, [2,18].DelayTimerSP := 1, [2,18].Priority := 1, [2,18].ActiveStateCFg := 1, [2,18].RealInputCfg := 1, [2,18].InputAddressCfg := 18, [2,18].OverrideCfg := 1, [2,18].PriorityCfg := 1, [2,19].AlarmCurrentValue := 1, [2,19].Override := 1, [2,19].DelayTimer.PRE := 1000, [2,19].DelayTimer.ACC := 1019, [2,19].DelayTimer.EN := 1, [2,19].DelayTimer.DN := 1, [2,19].DelayTimerSP := 1, [2,19].ActiveStateCFg := 1, [2,19].RealInputCfg := 1, [2,19].InputAddressCfg := 19, [2,19].OverrideCfg := 1, [2,19].PriorityCfg := 1, [2,20].AlarmCurrentValue := 1, [2,20].Override := 1, [2,20].DelayTimer.PRE := 1000,
        [2,20].DelayTimer.ACC := 1019, [2,20].DelayTimer.EN := 1, [2,20].DelayTimer.DN := 1, [2,20].DelayTimerSP := 1, [2,20].ActiveStateCFg := 1, [2,20].RealInputCfg := 1, [2,20].InputAddressCfg := 20, [2,20].OverrideCfg := 1, [2,20].PriorityCfg := 1, [2,21].AlarmCurrentValue := 1, [2,21].AlarmAck := 1, [2,21].Alarm := 1, [2,21].Mimic := 5, [2,21].DelayTimer.PRE := 1000, [2,21].DelayTimer.ACC := 1003, [2,21].DelayTimer.EN := 1, [2,21].DelayTimer.DN := 1, [2,21].DelayTimerSP := 1, [2,21].Priority := 1, [2,21].ActiveStateCFg := 1, [2,21].RealInputCfg := 1, [2,21].InputAddressCfg := 21, [2,21].AlarmONS := 1, [2,22].AlarmCurrentValue := 1, [2,22].AlarmAck := 1, [2,22].Alarm := 1, [2,22].Mimic := 5, [2,22].DelayTimer.PRE := 1000, [2,22].DelayTimer.ACC := 1004, [2,22].DelayTimer.EN := 1, [2,22].DelayTimer.DN := 1, [2,22].DelayTimerSP := 1, [2,22].Priority := 1, [2,22].ActiveStateCFg := 1, [2,22].RealInputCfg := 1, [2,22].InputAddressCfg := 22, [2,22].AlarmONS := 1, [2,23].AlarmCurrentValue := 1, [2,23].Override := 1, [2,23].DelayTimer.PRE := 1000, [2,23].DelayTimer.ACC := 1018, [2,23].DelayTimer.EN := 1, [2,23].DelayTimer.DN := 1, [2,23].DelayTimerSP := 1, [2,23].Priority := 1, [2,23].ActiveStateCFg := 1, [2,23].RealInputCfg := 1, [2,23].InputAddressCfg := 23, [2,23].OverrideCfg := 1, [2,23].PriorityCfg := 1, [2,24].AlarmCurrentValue := 1, [2,24].Override := 1, [2,24].DelayTimer.PRE := 1000, [2,24].DelayTimer.ACC := 1018, [2,24].DelayTimer.EN := 1, [2,24].DelayTimer.DN := 1, [2,24].DelayTimerSP := 1, [2,24].Priority := 1, [2,24].ActiveStateCFg := 1, [2,24].RealInputCfg := 1,
        [2,24].InputAddressCfg := 24, [2,24].OverrideCfg := 1, [2,24].PriorityCfg := 1, [2,25].AlarmCurrentValue := 1, [2,25].Override := 1, [2,25].DelayTimer.PRE := 20000, [2,25].DelayTimerSP := 2, [2,25].Priority := 1, [2,25].ActiveStateCFg := 1, [2,25].RealInputCfg := 1, [2,25].InputAddressCfg := 25, [2,25].OverrideCfg := 1, [2,25].PriorityCfg := 1, [2,25].Cond1Cfg := 1, [2,27].SoftInput := 1, [2,28].SoftInput := 1, [2,29].SoftInput := 1, [2,30].SoftInput := 1, [2,34].Tag := 'DI1', [2,34].Override := 1, [2,34].SoftInput := 1, [2,34].ActiveStateCFg := 1, [2,34].RealInputCfg := 1, [2,34].InputAddressCfg := 34, [2,34].OverrideCfg := 1, [2,34].PriorityCfg := 1, [2,35].Tag := 'DI2', [2,35].Override := 1, [2,35].ActiveStateCFg := 1, [2,35].RealInputCfg := 1, [2,35].InputAddressCfg := 35, [2,35].OverrideCfg := 1, [2,35].PriorityCfg := 1, [2,36].Tag := 'DI3', [2,36].Override := 1, [2,36].SoftInput := 1, [2,36].ActiveStateCFg := 1, [2,36].RealInputCfg := 1, [2,36].InputAddressCfg := 36, [2,36].OverrideCfg := 1, [2,36].PriorityCfg := 1, [2,37].Tag := 'DI4', [2,37].Override := 1, [2,37].ActiveStateCFg := 1, [2,37].RealInputCfg := 1, [2,37].InputAddressCfg := 37, [2,37].OverrideCfg := 1, [2,37].PriorityCfg := 1, [2,38].Tag := 'DI5', [2,38].Override := 1, [2,38].ActiveStateCFg := 1, [2,38].RealInputCfg := 1, [2,38].InputAddressCfg := 38, [2,38].OverrideCfg := 1, [2,38].PriorityCfg := 1, [2,39].Tag := 'DI6', [2,39].Override := 1, [2,39].SoftInput := 1, [2,39].ActiveStateCFg := 1, [2,39].RealInputCfg := 1,
        [2,39].InputAddressCfg := 39, [2,39].OverrideCfg := 1, [2,39].PriorityCfg := 1, [2,40].Tag := 'DI7', [2,40].Override := 1, [2,40].ActiveStateCFg := 1, [2,40].RealInputCfg := 1, [2,40].InputAddressCfg := 40, [2,40].OverrideCfg := 1, [2,40].PriorityCfg := 1, [2,41].Tag := 'DI8', [2,41].Override := 1, [2,41].SoftInput := 1, [2,41].ActiveStateCFg := 1, [2,41].RealInputCfg := 1, [2,41].InputAddressCfg := 41, [2,41].OverrideCfg := 1, [2,41].PriorityCfg := 1, [2,50].Tag := 'YA01', [2,50].AlarmCurrentValue := 1, [2,50].Alarm := 1, [2,50].Mimic := 2, [2,50].SoftInput := 1, [2,50].Condition1 := 1, [2,50].DelayTimer.PRE := 60000, [2,50].DelayTimer.ACC := 212, [2,50].DelayTimer.EN := 1, [2,50].DelayTimer.TT := 1, [2,50].DelayTimerSP := 60, [2,50].EnableCfg := 1, [2,50].InputAddressCfg := 50, [2,50].AlarmCfg := 1, [2,50].AlarmStateCfg := 1, [2,50].OverrideCfg := 1, [2,50].PriorityCfg := 1, [2,50].Cond1Cfg := 1, [2,50].AlarmONS := 1, [2,51].Tag := 'YA02', [2,51].AlarmCurrentValue := 1, [2,51].Alarm := 1, [2,51].Mimic := 2, [2,51].SoftInput := 1, [2,51].Condition1 := 1, [2,51].DelayTimer.PRE := 60000, [2,51].DelayTimer.ACC := 60018, [2,51].DelayTimer.EN := 1, [2,51].DelayTimer.DN := 1, [2,51].DelayTimerSP := 60, [2,51].EnableCfg := 1, [2,51].InputAddressCfg := 51, [2,51].AlarmCfg := 1, [2,51].AlarmStateCfg := 1, [2,51].OverrideCfg := 1, [2,51].PriorityCfg := 1, [2,51].Cond1Cfg := 1, [2,51].AlarmONS := 1, [2,52].Tag := 'YA03', [2,52].AlarmCurrentValue := 1, [2,52].Alarm := 1, [2,52].Mimic := 2,
        [2,52].SoftInput := 1, [2,52].Condition1 := 1, [2,52].DelayTimer.PRE := 60000, [2,52].DelayTimer.ACC := 4922, [2,52].DelayTimer.EN := 1, [2,52].DelayTimer.TT := 1, [2,52].DelayTimerSP := 60, [2,52].EnableCfg := 1, [2,52].InputAddressCfg := 52, [2,52].AlarmCfg := 1, [2,52].AlarmStateCfg := 1, [2,52].OverrideCfg := 1, [2,52].PriorityCfg := 1, [2,52].Cond1Cfg := 1, [2,52].AlarmONS := 1, [2,53].Tag := 'YA04', [2,53].DelayTimer.PRE := 60000, [2,53].DelayTimerSP := 60, [2,53].EnableCfg := 1, [2,53].ActiveStateCFg := 1, [2,53].InputAddressCfg := 53, [2,53].AlarmCfg := 1, [2,53].AlarmStateCfg := 1, [2,53].OverrideCfg := 1, [2,53].PriorityCfg := 1, [2,54].Tag := 'YA05', [2,54].DelayTimer.PRE := 60000, [2,54].DelayTimerSP := 60, [2,54].EnableCfg := 1, [2,54].ActiveStateCFg := 1, [2,54].InputAddressCfg := 54, [2,54].AlarmCfg := 1, [2,54].AlarmStateCfg := 1, [2,54].OverrideCfg := 1, [2,54].PriorityCfg := 1, [2,55].Tag := 'YA06', [2,55].CurrentValue := 1, [2,55].AlarmCurrentValue := 1, [2,55].AlarmAck := 1, [2,55].Alarm := 1, [2,55].Mimic := 5, [2,55].SoftInput := 1, [2,55].DelayTimer.PRE := 5000, [2,55].DelayTimer.ACC := 5022, [2,55].DelayTimer.EN := 1, [2,55].DelayTimer.DN := 1, [2,55].DelayTimerSP := 5, [2,55].Priority := 1, [2,55].EnableCfg := 1, [2,55].ActiveStateCFg := 1, [2,55].InputAddressCfg := 55, [2,55].AlarmCfg := 1, [2,55].AlarmStateCfg := 1, [2,55].OverrideCfg := 1, [2,55].PriorityCfg := 1, [2,55].AlarmONS := 1, [2,56].Tag := 'YA07', [2,56].DelayTimer.PRE := 2000, [2,56].DelayTimerSP := 2, [2,56].EnableCfg := 1,
        [2,56].ActiveStateCFg := 1, [2,56].InputAddressCfg := 56, [2,56].AlarmCfg := 1, [2,56].AlarmStateCfg := 1, [2,56].OverrideCfg := 1, [2,56].PriorityCfg := 1, [2,57].Tag := 'YA08', [2,57].CurrentValue := 1, [2,57].AlarmCurrentValue := 1, [2,57].AlarmAck := 1, [2,57].Alarm := 1, [2,57].Mimic := 5, [2,57].SoftInput := 1, [2,57].DelayTimer.PRE := 5000, [2,57].DelayTimer.ACC := 5023, [2,57].DelayTimer.EN := 1, [2,57].DelayTimer.DN := 1, [2,57].DelayTimerSP := 5, [2,57].Priority := 1, [2,57].EnableCfg := 1, [2,57].ActiveStateCFg := 1, [2,57].InputAddressCfg := 57, [2,57].AlarmCfg := 1, [2,57].AlarmStateCfg := 1, [2,57].OverrideCfg := 1, [2,57].PriorityCfg := 1, [2,57].AlarmONS := 1, [2,58].Tag := 'YA09', [2,58].DelayTimer.PRE := 2000, [2,58].DelayTimerSP := 2, [2,58].EnableCfg := 1, [2,58].ActiveStateCFg := 1, [2,58].InputAddressCfg := 58, [2,58].AlarmCfg := 1, [2,58].AlarmStateCfg := 1, [2,58].OverrideCfg := 1, [2,58].PriorityCfg := 1, [2,59].Tag := 'YA10', [2,59].CurrentValue := 1, [2,59].Mimic := 1, [2,59].Priority := 1, [2,59].EnableCfg := 1, [2,59].InputAddressCfg := 59, [2,59].AlarmCfg := 1, [2,59].AlarmStateCfg := 1, [2,60].Tag := 'YA11', [2,60].Override := 1, [2,60].DelayTimer.PRE := 5000, [2,60].DelayTimerSP := 5, [2,60].EnableCfg := 1, [2,60].ActiveStateCFg := 1, [2,60].InputAddressCfg := 60, [2,60].AlarmCfg := 1, [2,60].AlarmStateCfg := 1, [2,60].OverrideCfg := 1, [2,60].PriorityCfg := 1, [2,61].Tag := 'YA12', [2,61].EnableCfg := 1, [2,61].ActiveStateCFg := 1, [2,61].InputAddressCfg := 61,
        [2,61].AlarmCfg := 1, [2,61].AlarmStateCfg := 1, [2,61].OverrideCfg := 1, [2,61].PriorityCfg := 1, [2,62].Tag := 'YA13', [2,62].DelayTimer.PRE := 2000, [2,62].DelayTimerSP := 2, [2,62].EnableCfg := 1, [2,62].ActiveStateCFg := 1, [2,62].InputAddressCfg := 62, [2,62].AlarmCfg := 1, [2,62].AlarmStateCfg := 1, [2,62].OverrideCfg := 1, [2,62].PriorityCfg := 1, [2,63].Tag := 'YA14', [2,63].CurrentValue := 1, [2,63].Mimic := 1, [2,63].DelayTimer.PRE := 60000, [2,63].DelayTimerSP := 60, [2,63].EnableCfg := 1, [2,63].InputAddressCfg := 63, [2,63].AlarmCfg := 1, [2,63].AlarmStateCfg := 1, [2,64].Tag := 'UserNCr1', [2,64].CurrentValue := 1, [2,64].Mimic := 1, [2,64].EnableCfg := 1, [2,64].InputAddressCfg := 64, [2,65].Tag := 'UserCr1', [2,65].CurrentValue := 1, [2,65].Mimic := 1, [2,65].Priority := 1, [2,65].EnableCfg := 1, [2,65].InputAddressCfg := 65, [2,66].Tag := 'UserNCr2', [2,66].CurrentValue := 1, [2,66].Mimic := 1, [2,66].DelayTimer.PRE := 2000, [2,66].DelayTimerSP := 2, [2,66].EnableCfg := 1, [2,66].InputAddressCfg := 66, [2,67].Tag := 'UserCr2', [2,67].CurrentValue := 1, [2,67].Mimic := 1, [2,67].DelayTimer.PRE := 2000, [2,67].DelayTimerSP := 2, [2,67].Priority := 1, [2,67].EnableCfg := 1, [2,67].InputAddressCfg := 67, [2,68].Tag := 'ZSDF', [2,68].CurrentValue := 1, [2,68].AlarmCurrentValue := 1, [2,68].AlarmAck := 1, [2,68].Alarm := 1, [2,68].Mimic := 5, [2,68].SoftInput := 1, [2,68].DelayTimer.PRE := 1000, [2,68].DelayTimer.ACC := 1042, [2,68].DelayTimer.EN := 1, [2,68].DelayTimer.DN := 1,
        [2,68].DelayTimerSP := 1, [2,68].Priority := 1, [2,68].EnableCfg := 1, [2,68].ActiveStateCFg := 1, [2,68].InputAddressCfg := 68, [2,68].AlarmCfg := 1, [2,68].AlarmStateCfg := 1, [2,68].OverrideCfg := 1, [2,68].PriorityCfg := 1, [2,68].AlarmONS := 1, [2,69].Tag := 'YA15', [2,69].CurrentValue := 1, [2,69].AlarmCurrentValue := 1, [2,69].AlarmAck := 1, [2,69].Alarm := 1, [2,69].Mimic := 5, [2,69].SoftInput := 1, [2,69].DelayTimer.PRE := 5000, [2,69].DelayTimer.ACC := 2039, [2,69].DelayTimer.EN := 1, [2,69].DelayTimer.DN := 1, [2,69].DelayTimerSP := 5, [2,69].Priority := 1, [2,69].EnableCfg := 1, [2,69].ActiveStateCFg := 1, [2,69].InputAddressCfg := 69, [2,69].AlarmCfg := 1, [2,69].AlarmStateCfg := 1, [2,69].OverrideCfg := 1, [2,69].PriorityCfg := 1, [2,69].AlarmONS := 1, [2,70].Tag := 'YA16', [2,70].DelayTimer.PRE := 2000, [2,70].DelayTimerSP := 2, [2,70].EnableCfg := 1, [2,70].ActiveStateCFg := 1, [2,70].InputAddressCfg := 70, [2,70].AlarmCfg := 1, [2,70].AlarmStateCfg := 1, [2,70].OverrideCfg := 1, [2,70].PriorityCfg := 1, [2,71].Tag := 'YA17', [2,71].CurrentValue := 1, [2,71].AlarmCurrentValue := 1, [2,71].AlarmAck := 1, [2,71].Alarm := 1, [2,71].Mimic := 5, [2,71].SoftInput := 1, [2,71].DelayTimer.PRE := 5000, [2,71].DelayTimer.ACC := 2036, [2,71].DelayTimer.EN := 1, [2,71].DelayTimer.DN := 1, [2,71].DelayTimerSP := 5, [2,71].Priority := 1, [2,71].EnableCfg := 1, [2,71].ActiveStateCFg := 1, [2,71].InputAddressCfg := 71, [2,71].AlarmCfg := 1, [2,71].AlarmStateCfg := 1, [2,71].OverrideCfg := 1,
        [2,71].PriorityCfg := 1, [2,71].AlarmONS := 1, [2,72].Tag := 'YA18', [2,72].DelayTimer.PRE := 2000, [2,72].DelayTimerSP := 2, [2,72].EnableCfg := 1, [2,72].ActiveStateCFg := 1, [2,72].InputAddressCfg := 72, [2,72].AlarmCfg := 1, [2,72].AlarmStateCfg := 1, [2,72].OverrideCfg := 1, [2,72].PriorityCfg := 1, [2,73].Tag := 'YA19', [2,73].CurrentValue := 1, [2,73].AlarmCurrentValue := 1, [2,73].AlarmAck := 1, [2,73].Alarm := 1, [2,73].Mimic := 5, [2,73].SoftInput := 1, [2,73].DelayTimer.PRE := 5000, [2,73].DelayTimer.ACC := 2036, [2,73].DelayTimer.EN := 1, [2,73].DelayTimer.DN := 1, [2,73].DelayTimerSP := 5, [2,73].Priority := 1, [2,73].EnableCfg := 1, [2,73].ActiveStateCFg := 1, [2,73].InputAddressCfg := 73, [2,73].AlarmCfg := 1, [2,73].AlarmStateCfg := 1, [2,73].OverrideCfg := 1, [2,73].PriorityCfg := 1, [2,73].AlarmONS := 1, [2,74].Tag := 'YA20', [2,74].DelayTimer.PRE := 2000, [2,74].DelayTimerSP := 2, [2,74].EnableCfg := 1, [2,74].ActiveStateCFg := 1, [2,74].InputAddressCfg := 74, [2,74].AlarmCfg := 1, [2,74].AlarmStateCfg := 1, [2,74].OverrideCfg := 1, [2,74].PriorityCfg := 1, [2,75].Tag := 'YA21', [2,75].CurrentValue := 1, [2,75].AlarmCurrentValue := 1, [2,75].AlarmAck := 1, [2,75].Alarm := 1, [2,75].Mimic := 5, [2,75].SoftInput := 1, [2,75].DelayTimer.PRE := 5000, [2,75].DelayTimer.ACC := 2036, [2,75].DelayTimer.EN := 1, [2,75].DelayTimer.DN := 1, [2,75].DelayTimerSP := 5, [2,75].Priority := 1, [2,75].EnableCfg := 1, [2,75].ActiveStateCFg := 1, [2,75].InputAddressCfg := 75, [2,75].AlarmCfg := 1,
